(* IEC 61131-3 sources: daoli-st-library/DL_MathData (part 6) *)

(* ---- FC_DL_StringToUdintEx.st ---- *)
(*
    组件名称 : FC_DL_StringToUdintEx
    所属子库 : DL_MathData
    当前版本 : 1.0.0
    兼 容 性 : CODESYS V3.5+ / TwinCAT 3 / 汇川 InoProShop；仅依赖 Standard.library
    溯源声明 : IEC 61131-3 标准语义的道莅防御性实现
              （解析口径复用库内 FC_DL_StringToDint 的四态状态机与判界结构，
                按无符号域重写判界；零外部源码复制，参考实现仅限 MIT/Apache 许可）
    功能描述 : 无符号整数字符串严格解析（UDINT 域，配方号 / 计数器预置 / 批次号）。
              取舍 ①：不委托任何平台串转数值内建——三家平台对非法字符、前导空格、
              符号重复的处理各不相同，有的返回 0、有的抛异常、有的静默截断，且都
              不告诉调用方错在第几位；本件逐字符推进，判断口径完全一致，并给出
              首个非法字符位置。
              取舍 ②：空格一律按非法字符拒绝（与 FC_DL_StringToDint 的「忽略空格
              并提示」口径刻意分叉）——UDINT 域多为机器写入值，隐式吞空格易掩盖
              脏数据，从严拒绝并在 nErrPos 定位。
              取舍 ③：升位到 LINT 累加，每步先判界再落账——UDINT 域中间量在
              429496729 × 10 + 5 处已越界，直接在 UDINT/DINT 里累加必然回绕
              （R241 口径：跨类型降型禁靠隐式回绕兜底）；LINT 域足够宽，判界
              判的是 LINT 与 UDINT 上界的比较，安全。
              取舍 ④：溢出后返回「夹到上界」的值并置 bValid = FALSE——夹域值便于
              现场看出「方向对了但超了」；同时绝不把夹域值当有效值输出。
              取舍 ⑤：负号一律判越域拒绝（含 −0）——UDINT 无负域，负号属语义错误
              而非语法错误，独立占码与非法字符区分。
    本文件内含 : FUNCTION FC_DL_StringToUdintEx（单 POU）
                 同文件 TYPE E_DL_StrToUdintState（归属本函数，全库唯一）
    依 赖    : 无 DL_ 内部依赖；Standard.library: LEN / MID / FIND
    错误码   : 16#0001_03D6 [故障级] 空串或仅符号，nErrPos = 长度 + 1，返回 0，bValid = FALSE
               16#0001_03D7 [故障级] 负值越 UDINT 域（含 −0，从严拒绝），返回 0，bValid = FALSE
               16#0001_03D8 [故障级] 数值溢出，返回夹到上界的值，bValid = FALSE
               16#0001_03D9 [故障级] 非法字符（含 CASE 落 ELSE 的非法状态兜底与扫描失控复用，
                             不新占码位），返回 0，bValid = FALSE
               （R90 反证句：四类故障场景的输出组合互不相同——空串与非法字符返回 0、
                 溢出返回上界夹域值、负值返回 0 但 nErrPos 定位在符号位；返回值加
                 nErrPos 无法唯一还原「空串」与「负值」（同为 0），故两场景各自占码）
    红线自检 : R1 ✓ 零全局变量与外部变量 ｜ R2 ✓ 零物理 IO 地址
              R3 ✓ 纯 IEC 61131-3 ｜ R4 ✓ 空串闸 + 非法字符定位 + 先判界后落账 + WHILE 守卫计数器
              R5 ✓ 全变量中英双语同行注释 ｜ R6 ✓ ENUM + CASE + ELSE 兜底（非法状态复用 03D9）
              R7 N/A 无定时器、无沿检测实例 ｜ R8 ✓ 上下界、长度上限、守卫上限全常量化
    修订历史 :
        2026-11-19  v1.0.0  首版，R40 批次 3 入库
*)

(*-----------------------------------------------------------------------------
 * 枚举: E_DL_StrToUdintState（归属本函数，与其同文件发布，全库唯一）
 * 含义: 逐字符解析的四态推进，成员值写死便于工程持久化
 *----------------------------------------------------------------------------*)
TYPE E_DL_StrToUdintState :
(
    eLeadSpace := 0,    // 起始态：空格按非法字符拒绝，遇其余字符转符号态 ｜ start state, blanks are rejected as illegal, any other character moves to the sign state
    eSign      := 10,   // 符号态：取前导 +/− 号或直接进数字态 ｜ sign state, consumes the leading sign or falls through to the digits
    eDigits    := 20,   // 数字态：逐位累加，遇非数字一律非法 ｜ digits state, accumulates digit by digit, any non-digit is illegal
    eDone      := 30    // 结束态：串尾守卫态，任何字符均非法 ｜ done state, an end-of-string guard, any character here is illegal
);
END_TYPE

FUNCTION FC_DL_StringToUdintEx : UDINT
VAR_INPUT
    sIn             : STRING;           // 待解析文本，最长 255 字符，不允许任何空格 [字符] ｜ input text, up to 255 characters, no blanks allowed [char]
    bAllowSign      : BOOL := FALSE;    // 是否允许前导 +/− 号，UDINT 口径缺省禁止 ｜ whether a leading sign is allowed, the UDINT mode forbids it by default
END_VAR
VAR_OUTPUT
    eErr            : UDINT;           // 错误码，0=正常；16#0001_03XX 故障级 ｜ error id, 0=ok, 16#0001_03XX=fault level
    bError          : BOOL;            // 故障级标志，eErr 落 16#0001_03XX 时为 TRUE ｜ fault flag, TRUE on fault-level eErr
    bValid          : BOOL;            // 返回值是否可用 ｜ result usable flag
    nErrPos         : INT;             // 首个非法字符位置（1 基），0 = 无错 [字符] ｜ position of the first illegal character, 1 based, zero means no error [char]
END_VAR
VAR
    eState          : E_DL_StrToUdintState;  // 解析状态机当前态 ｜ current parse state
    nLen            : INT;             // 文本长度，入口锁存一次，其后全部取自该副本 [字符] ｜ latched text length, every later bound comes from this copy [char]
    nPos            : INT;             // 字符游标（1 基）[字符] ｜ character cursor, 1 based [char]
    nGuard          : DINT;            // WHILE 防死锁守卫计数 [次] ｜ loop guard counter [count]
    nDigitVal       : INT;             // 当前字符的数字值，未命中为 −1 [无量纲] ｜ numeric value of the current character, minus one when not a digit [dimensionless]
    nDigits         : INT;             // 已接受的有效数字位数 [位] ｜ number of accepted digits [digit]
    sChar           : STRING(1);       // 当前字符，由标准 MID 取出 [字符] ｜ current character read with the standard MID [char]
    bNeg            : BOOL;            // 负号标志，由前导符号决定 ｜ negative flag set by the leading sign
    bAbort          : BOOL;            // 中止标志，置位后立即退出扫描 ｜ abort flag, the scan stops as soon as it is set
    bOverflow       : BOOL;            // 溢出标志 ｜ overflow flag
    liAcc           : LINT;            // 升位累加器 [无量纲] ｜ widened accumulator [dimensionless]
    liNext          : LINT;            // 下一拍候选累加值，先判界再落账 [无量纲] ｜ candidate accumulator tested before it is committed [dimensionless]
END_VAR
VAR CONSTANT
    DL_UDINT_MAX_LI    : LINT := 4294967295;     // UDINT 上界的 LINT 判界值 [无量纲] ｜ UDINT upper bound as the LINT test limit [dimensionless]
    DL_LINT_TEN        : LINT := 10;             // 十进制进位基数 [无量纲] ｜ decimal radix [dimensionless]
    DL_STR_MAXLEN      : INT := 255;             // 文本长度上限 [字符] ｜ text length upper bound [char]
    DL_STR_GUARD_MAX   : DINT := 600;            // 守卫上限，须大于 255 + 2 次不推进状态 ｜ guard limit, larger than the length plus two non advancing states
    DL_STR_ONE         : INT := 1;               // 单位哨兵 [无量纲] ｜ unity sentinel [dimensionless]
    DL_STR_DIGITS      : STRING := '0123456789'; // 数字字符表，FIND 命中位置 − 1 即数字值 [字符] ｜ digit table, the FIND position minus one is the value [char]
    DL_ERR_NONE        : UDINT := 16#0000_0000;  // 无故障 ｜ no error
END_VAR

// 段 1｜返回值与错误状态预置 ｜ segment 1, preset the return value and the error state
FC_DL_StringToUdintEx := 0;                   // 故障缺省返回 0 ｜ fault default returns zero
eErr           := DL_ERR_NONE;                // 预置无错误 ｜ preset no error
bError         := FALSE;                      // 预置无故障 ｜ preset no fault
bValid         := FALSE;                      // 预置结果不可用 ｜ preset unusable
nErrPos        := 0;                          // 0 表示无错 ｜ zero means no error
eState         := E_DL_StrToUdintState.eLeadSpace;  // 起始态 ｜ start in the start state
nLen           := LEN(sIn);                   // 长度只锁存一次，禁循环内重复 LEN ｜ latch the length once, never call LEN again in the loop
nPos           := DL_STR_ONE;                 // 游标从 1 开始（MID 为 1 基）｜ the cursor starts at one because MID is one based
nGuard         := 0;                          // 守卫清零 ｜ clear the guard
nDigits        := 0;                          // 有效位数清零 ｜ clear the digit count
nDigitVal      := 0;                          // 数字值清零 ｜ clear the digit value
bNeg           := FALSE;                      // 预置无负号 ｜ preset no negative sign
bAbort         := FALSE;                      // 预置不中止 ｜ preset no abort
bOverflow      := FALSE;                      // 预置无溢出 ｜ preset no overflow
liAcc          := 0;                          // 累加器清零 ｜ clear the accumulator
liNext         := 0;                          // 候选值清零 ｜ clear the candidate
sChar          := '';                         // 字符缓冲清空 ｜ clear the character buffer

// 段 2｜逐字符状态机：四态推进，ELSE 兜底拦非法状态 ｜ segment 2, four state machine with an ELSE backstop
WHILE (nPos <= nLen) AND (NOT bAbort) AND (nGuard <= DL_STR_GUARD_MAX) DO
    sChar := MID(sIn, DL_STR_ONE, nPos);    // 取当前位置的一个字符 ｜ take one character at the current position
    CASE eState OF
        E_DL_StrToUdintState.eLeadSpace :
            // 起始态：空格从严拒绝（取舍 ②），其余字符转符号态 ｜ start state: blanks are strictly rejected, any other character moves to the sign state
            IF sChar = ' ' THEN
                eErr    := 16#0001_03D9;    // 空格按非法字符拒绝（故障级）｜ a blank is rejected as an illegal character
                bError  := TRUE;            // 置故障标志 ｜ raise the fault flag
                nErrPos := nPos;            // 定位到空格位 ｜ point at the blank
                bAbort  := TRUE;            // 中止扫描 ｜ abort the scan
            ELSE
                eState := E_DL_StrToUdintState.eSign;  // 转符号态，本拍不消费字符，下一轮重取同一字符 ｜ move to the sign state without consuming this character
            END_IF

        E_DL_StrToUdintState.eSign :
            IF (sChar = '+') OR (sChar = '-') THEN
                IF NOT bAllowSign THEN
                    eErr   := 16#0001_03D9;     // 不允许符号却出现符号（故障级）｜ a sign appeared although it is forbidden
                    bError := TRUE;             // 置故障标志 ｜ raise the fault flag
                    nErrPos := nPos;            // 定位到符号位 ｜ point at the sign
                    bAbort := TRUE;             // 中止扫描 ｜ abort the scan
                ELSE
                    bNeg   := (sChar = '-');    // 负号判定（取舍 ⑤：负号在出口判越域）｜ detect the minus sign (rejected as out-of-domain at the exit)
                    nPos   := nPos + DL_STR_ONE;   // 消费符号 ｜ consume the sign
                    eState := E_DL_StrToUdintState.eDigits;  // 转数字态 ｜ move to the digit state
                END_IF
            ELSE
                eState := E_DL_StrToUdintState.eDigits;  // 无符号直接进数字态 ｜ no sign, go straight to the digits
            END_IF

        E_DL_StrToUdintState.eDigits :
            // 数字态：数字先判界后落账，非数字一律非法（空格含在内，从严口径）｜ digit state: digits are tested before commit, any non-digit is illegal (blanks included, strict mode)
            nDigitVal := FIND(DL_STR_DIGITS, sChar) - DL_STR_ONE;   // 命中 0~9，未命中 −1 ｜ zero to nine when found, minus one otherwise
            IF nDigitVal < 0 THEN
                eErr    := 16#0001_03D9;            // 非法字符（故障级）｜ illegal character, fault level
                bError  := TRUE;                    // 置故障标志 ｜ raise the fault flag
                nErrPos := nPos;                    // 定位到首个非法字符 ｜ point at the first illegal character
                bAbort  := TRUE;                    // 中止扫描 ｜ abort the scan
            ELSE
                liNext := liAcc * DL_LINT_TEN + INT_TO_LINT(nDigitVal);   // 先算候选值 ｜ compute the candidate first
                IF liNext > DL_UDINT_MAX_LI THEN
                    bOverflow := TRUE;              // 越界即溢出，不落账 ｜ beyond the limit means overflow, not committed
                    nErrPos   := nPos;              // 溢出位也必须定位，否则 nErrPos = 0 会被读成「无错」｜ locate the overflowing digit, zero would read as no error
                    bAbort    := TRUE;              // 中止扫描 ｜ abort the scan
                ELSE
                    liAcc   := liNext;              // 落账 ｜ commit
                    nDigits := nDigits + DL_STR_ONE;   // 有效位加一 ｜ one more digit accepted
                    nPos    := nPos + DL_STR_ONE;   // 前进一格 ｜ advance one position
                END_IF
                IF nPos > nLen THEN
                    eState := E_DL_StrToUdintState.eDone;   // 已到串尾，转结束态守卫 ｜ reached the end, move to the done guard
                END_IF
            END_IF

        E_DL_StrToUdintState.eDone :
            // 结束态：本件从严口径，任何尾随字符（含空格）均非法 ｜ done state: in strict mode any trailing character (blanks included) is illegal
            eErr    := 16#0001_03D9;                // 尾随非法字符（故障级）｜ illegal trailing character, fault level
            bError  := TRUE;                        // 置故障标志 ｜ raise the fault flag
            nErrPos := nPos;                        // 定位 ｜ point at the position
            bAbort  := TRUE;                        // 中止扫描 ｜ abort the scan

    ELSE
        // 非法状态兜底：枚举被外部改写或内存损伤，一律按「输入不可解析」处置（R90：复用非法字符码，不新占码位）
        eState   := E_DL_StrToUdintState.eDone;          // 强制回已知态 ｜ force back to a known state
        eErr     := 16#0001_03D9;                        // 复用非法字符码 ｜ reuse the illegal character code
        bError   := TRUE;                               // 置故障标志 ｜ raise the fault flag
        nErrPos  := nPos;                               // 定位当前位 ｜ point at the current position
        bAbort   := TRUE;                               // 中止扫描 ｜ abort the scan
    END_CASE
    nGuard := nGuard + 1;                              // 守卫递增 ｜ increment the guard
END_WHILE

// 段 3｜守卫复检：理论不可达（长度 ≤ 255，不推进状态最多 2 次）｜ segment 3, guard re-check, unreachable in theory
IF nGuard > DL_STR_GUARD_MAX THEN
    FC_DL_StringToUdintEx := 0;        // 不给可疑结果 ｜ never emit a suspicious result
    eErr   := 16#0001_03D9;            // 扫描失控复用非法字符码（不新占码位）｜ a runaway scan reuses the illegal character code
    bError := TRUE;                    // 置故障标志 ｜ raise the fault flag
    nErrPos := nPos;                   // 定位 ｜ point at the current position
    RETURN;                            // bValid 保持 FALSE ｜ bValid stays FALSE
END_IF

// 段 4｜非法/溢出已中止：直接出口（故障行为已在扫描中定性）｜ segment 4, exit when the scan was aborted
IF bAbort THEN
    IF bOverflow THEN
        FC_DL_StringToUdintEx := 4294967295; // 溢出夹到 UDINT 上界 ｜ overflow saturated to the UDINT upper bound
        eErr := 16#0001_03D8;        // 溢出已夹上界（故障级）｜ overflow saturated, fault level
        bError := TRUE;              // 置故障标志（R45 配对，扫描内溢出只置 bOverflow，出口统一配对）｜ raise the fault flag (R45 pairing)
    ELSE
        FC_DL_StringToUdintEx := 0;  // 语法错误返回 0 ｜ a syntax error returns zero
    END_IF
    RETURN;                          // bValid 保持 FALSE ｜ bValid stays FALSE
END_IF

// 段 5｜空串或仅符号闸 ｜ segment 5, empty string or sign-only gate
IF nDigits = 0 THEN
    FC_DL_StringToUdintEx := 0;         // 无有效数字返回 0 ｜ no digit at all, return zero
    eErr    := 16#0001_03D6;            // 空串或仅符号（故障级）｜ empty or sign only, fault level
    bError  := TRUE;                    // 置故障标志（R45 配对）｜ raise the fault flag (R45 pairing)
    nErrPos := nLen + DL_STR_ONE;       // 指向「串尾后一位」，与库内同族口径一致 ｜ point past the end, consistent with the sibling component
    RETURN;                             // bValid 保持 FALSE ｜ bValid stays FALSE
END_IF

// 段 6｜负值越域闸（取舍 ⑤：负号含 −0 一律从严拒绝）｜ segment 6, negative out-of-domain gate (a minus sign including minus zero is strictly rejected)
IF bNeg THEN
    FC_DL_StringToUdintEx := 0;         // 负值越域返回 0 ｜ out-of-domain negative returns zero
    eErr    := 16#0001_03D7;            // 负值越 UDINT 域（故障级）｜ negative beyond the UDINT domain, fault level
    bError  := TRUE;                    // 置故障标志（R45 配对）｜ raise the fault flag (R45 pairing)
    nErrPos := DL_STR_ONE;              // 定位到符号位（第 1 位）｜ point at the sign position (position one)
    RETURN;                             // bValid 保持 FALSE ｜ bValid stays FALSE
END_IF

// 段 7｜出口装配：累加器域内单点落账 ｜ segment 7, exit assembly: the accumulator is in-domain, commit once
FC_DL_StringToUdintEx := LINT_TO_UDINT(liAcc); // 判界已保证 liAcc ≤ UDINT 上界，降型安全 ｜ the domain test guarantees the accumulator is within the UDINT bound, the down-conversion is safe
bValid := TRUE;                      // 结果可用 ｜ the result is usable
END_FUNCTION

(* ---- FC_DL_SwapBytes32.st ---- *)
(*==============================================================================
 * 组件名称 (Component)  : FC_DL_SwapBytes32
 * 所属子库 (Sublibrary) : DL_MathData
 * 当前版本 (Version)    : 1.0.0
 * 兼容性   (Platform)   : CODESYS 3.5 / TwinCAT 3 / 汇川 InoProShop / Machine Expert
 *                         仅依赖 Standard.library 的 SHL / SHR / AND / OR，零厂商方言
 * 功能描述 (Function)   : 32 位量四排布（ABCD / DCBA / BADC / CDAB）归一化转换。
 *                         调用方声明通信侧原始拼接值实际所属的排布，
 *                         函数统一输出 ABCD（大端大字）归一化值。
 *                         语义锁定为单向归一化，不做双向目标排布选择；
 *                         需要反向时以对称排布重新声明即可（四排布两两互逆）。
 *                         用于 Modbus 多寄存器浮点/长整型量"读回 1e38 天文数字"的定位与校正。
 * 开源溯源 (Origin)     : 原创实现。四种排布命名与业界别名（字交换 / 寄存器内字节互换 /
 *                         全反序）参照 modbus.org 公开协议说明与多家转换器技术资料的
 *                         事实约定；本文件为独立重构，未复制任何源码。
 * 本文件内含       : TYPE  E_DL_ByteOrder（配套枚举，归属 DL_MathData）
 *                    FC    FC_DL_SwapBytes32
 * 依赖     (Depends)    : 无 DL_ 内部依赖；Standard.library: SHL / SHR
 * 红线自检 (Redline)    : R1 ✓ 禁用全局存储与物理寻址 ｜ R2 ✓ 无地址直写
 *                         R3 ✓ 移位掩码提取 + 显式类型转换，无切片/指针/字节方言
 *                         R4 N/A（无除法/数组/循环/浮点）｜ R5 ✓ 全变量中英双语同行注释
 *                         R6 ✓ 四排布 CASE 分派 + ELSE 兜底 ｜ R7 N/A（无定时器/边沿实例）
 *                         R8 ✓ 移位量与掩码全常量化
 *
 * 【实现选择 / Implementation choice（边界 B6）】
 *   四条转换路径全部用"移位提取 + 显式 BYTE 转换 + 移位重装"实现，
 *   不调用 16 位互换构件，保证本文件自洽、可单独编译与单独单测。
 *
 * 【浮点使用口径 / Float usage（边界 B7）】
 *   本函数只输出归一化 DWORD，不做 DWORD 到 REAL 的二进制重解释。
 *   浮点拼接规则各平台存在差异，由调用方按其平台口径完成，避免在本层引入行为分支。
 *
 * 【验收向量 / Acceptance vectors（边界 B5，已复算）】
 *   以 16#12345678 为基准：ABCD → 16#12345678；DCBA → 16#78563412；
 *   BADC → 16#34127856；CDAB → 16#56781234。
 *
 * 修订历史 (Revision)   :
 *   2026-11-14  v1.0.0  首版入库（Phase 1 第二轮 · Level 0 批次 C）
 *============================================================================*)

(*-----------------------------------------------------------------------------
 * 枚举: E_DL_ByteOrder（归属 DL_MathData，与 FC_DL_SwapBytes32 同文件）
 * 含义: 通信侧 32 位量的字节排布。A 为最高字节（位 31..24），D 为最低字节。
 *----------------------------------------------------------------------------*)
TYPE E_DL_ByteOrder :
(
    eAbcd := 0,    // ABCD：大端大字（Modicon 事实标准），原始值无需转换 / Big-endian big-word, pass-through
    eDcba := 1,    // DCBA：四字节全反序，常见于小端 CPU 直出的协议栈 / Full byte reverse
    eBadc := 2,    // BADC：两个寄存器内部各自字节互换 / Byte swap within each register
    eCdab := 3     // CDAB：高低字交换（寄存器字序反），常见于电能表 / Word swap
);
END_TYPE

FUNCTION FC_DL_SwapBytes32 : DWORD
VAR_INPUT
    uRaw      : DWORD;                        // 通信侧原始 32 位拼接值 / Raw 32-bit value assembled from comms
    eRawOrder : E_DL_ByteOrder := eAbcd;      // 声明原始值所属排布 / Declared byte order of raw value
END_VAR
VAR_OUTPUT
    bValid    : BOOL;                         // 排布枚举合法标志 / Order enum valid flag
    uErrorId  : UDINT;                        // 故障码，0 = 无故障 / Error code, 0 = no error
END_VAR
VAR
    uA : BYTE;   // 字节 A（uRaw 位 31..24） / Byte A, bits 31..24
    uB : BYTE;   // 字节 B（uRaw 位 23..16） / Byte B, bits 23..16
    uC : BYTE;   // 字节 C（uRaw 位 15..8）  / Byte C, bits 15..8
    uD : BYTE;   // 字节 D（uRaw 位 7..0）   / Byte D, bits 7..0
END_VAR
VAR CONSTANT
    DL_SWAP_SHIFT8  : UDINT := 8;               // 字节移位量 [bit] / Byte shift width [bit]
    DL_SWAP_SHIFT16 : UDINT := 16;              // 字移位量 [bit] / Word shift width [bit]
    DL_SWAP_SHIFT24 : UDINT := 24;              // 最高字节移位量 [bit] / Top byte shift width [bit]
    DL_MASK_BYTE    : DWORD := 16#0000_00FF;    // 单字节掩码 / Single-byte mask
END_VAR

(*------------------------------------------------------------------------------
 * 段 1｜安全预置（边界 B1 / P-01）：先返回原值，任何异常路径都不会返回 0
 *      Safe preset: return the raw value first, no exceptional path returns zero
 *      0 对浮点量是合法灾难值，原值直通是最安全的确定值
 *      Zero is a legal but catastrophic float value, pass-through is the safest result
 *-----------------------------------------------------------------------------*)
FC_DL_SwapBytes32 := uRaw;
bValid   := TRUE;
uErrorId := 16#0000_0000;

(*------------------------------------------------------------------------------
 * 段 2｜字节提取（边界 B2）：仅移位 + 掩码 + 显式 BYTE 转换，禁止切片与指针
 *      Byte extraction: shift + mask + explicit BYTE conversion only
 *-----------------------------------------------------------------------------*)
uA := DWORD_TO_BYTE(SHR(uRaw, DL_SWAP_SHIFT24) AND DL_MASK_BYTE);
uB := DWORD_TO_BYTE(SHR(uRaw, DL_SWAP_SHIFT16) AND DL_MASK_BYTE);
uC := DWORD_TO_BYTE(SHR(uRaw, DL_SWAP_SHIFT8)  AND DL_MASK_BYTE);
uD := DWORD_TO_BYTE(uRaw AND DL_MASK_BYTE);

(*------------------------------------------------------------------------------
 * 段 3｜四排布分派（边界 B3/B4）：CASE 分派禁止 IF 链，ELSE 兜底拒收非法枚举
 *      Four-order dispatch: CASE only, ELSE intercepts an out-of-domain enum
 *-----------------------------------------------------------------------------*)
CASE eRawOrder OF

    eAbcd:
        (* 大端大字已是归一化目标，原值直通 *)
        (* Big-endian big-word is already the normalised target, pass through *)
        FC_DL_SwapBytes32 := uRaw;

    eDcba:
        (* 全反序：D C B A *)
        (* Full byte reverse: D C B A *)
        FC_DL_SwapBytes32 := (SHL(BYTE_TO_DWORD(uD), DL_SWAP_SHIFT24)
                          OR  SHL(BYTE_TO_DWORD(uC), DL_SWAP_SHIFT16)
                          OR  SHL(BYTE_TO_DWORD(uB), DL_SWAP_SHIFT8)
                          OR  BYTE_TO_DWORD(uA));

    eBadc:
        (* 寄存器内字节互换：B A D C *)
        (* Byte swap within each register: B A D C *)
        FC_DL_SwapBytes32 := (SHL(BYTE_TO_DWORD(uB), DL_SWAP_SHIFT24)
                          OR  SHL(BYTE_TO_DWORD(uA), DL_SWAP_SHIFT16)
                          OR  SHL(BYTE_TO_DWORD(uD), DL_SWAP_SHIFT8)
                          OR  BYTE_TO_DWORD(uC));

    eCdab:
        (* 高低字交换：C D A B *)
        (* Word swap: C D A B *)
        FC_DL_SwapBytes32 := (SHL(BYTE_TO_DWORD(uC), DL_SWAP_SHIFT24)
                          OR  SHL(BYTE_TO_DWORD(uD), DL_SWAP_SHIFT16)
                          OR  SHL(BYTE_TO_DWORD(uA), DL_SWAP_SHIFT8)
                          OR  BYTE_TO_DWORD(uB));

    ELSE
        (* 非法枚举拦截：枚举被强制写入定义域外的值时返回原值并报错 *)
        (* Illegal enum interception: keep the raw value and raise the error *)
        FC_DL_SwapBytes32 := uRaw;
        bValid            := FALSE;
        uErrorId          := 16#0001_000E;

END_CASE;
END_FUNCTION

(* ---- FC_DL_TableIndexBinarySearch.st ---- *)
(*==============================================================================
 * 组件名称 (Component)  : FC_DL_TableIndexBinarySearch
 * 所属子库 (Sublibrary) : DL_MathData
 * 当前版本 (Version)    : 1.0.0
 * 兼容性   (Platform)   : CODESYS 3.5+ / TwinCAT 3 / 汇川 InoProShop / 施耐德 Machine Expert
 *                         仅依赖 IEC 61131-3 标准数学（ABS / MIN / MAX），零厂商私有库
 * 功能描述 (Function)   : **升序**节点表二分查找定位（O(log n)），返回区间左端下标与段内比例。
 *                         迭代式二分：维护 [iLo, iHi] 使 afX[iLo] <= fXin <= afX[iHi]，
 *                         每次收缩一半，直到 iHi - iLo = 1，此时 iSeg = iLo。
 *                         32 点表最多 5 次迭代（2^5 = 32），循环上界显式封顶 8 次，
 *                         结构上不可能死循环（R6 周期安全：纯函数虽无跨周期状态，
 *                         仍对不可终止循环做硬保护）。
 *                         用途：大表（温压补偿、阀门口径选型）的高频查表，替代线性扫描。
 * 接口     (Interface)  : 输入 afX 升序节点表 [任意工程量]、iCount 有效点数 [个]（2..32）、
 *                         fXin 查询点 [同 afX 单位]；
 *                         输出 iSeg 区间左端下标 [1..iCount-1]、fRatio 段内比例 [0..1]、
 *                         bExact 是否恰命中节点、bClamped 越界钳位回执、
 *                         eErrCode（E_DL_TblBsearchErr）；
 *                         返回值 = bValid 定位可信标志（TRUE = iSeg/fRatio 可信）。
 * 边界     (Boundary)   : ① 属主边界：只做定位，不做取值；表必须升序（降序表用
 *                         FC_DL_TableLookupDescending）。
 *                         ② 点数域闸 2..32；越域 → 故障级 eBadCount。
 *                         ③ 非有限双判：查询点 + 全部表元素逐项枚举（漏判单个元素会使比较静默失效）。
 *                         ④ 升序性校验：二分不校验全序，但会校验命中区间的两个端点是否满足
 *                         afX[iSeg] <= afX[iSeg+1]，违反即判 eTableNotAsc（防止强序假设）。
 *                         ⑤ 段宽近似零 → fRatio 置 0 并置信息级 eDegenerateSeg（除零防护）。
 *                         ⑥ 迭代次数硬上界 DL_TBC_ITER_MAX = 8，超出即判 eSearchOverflow
 *                         （理论上不可达，作为不可终止循环的兜底闸）。
 *                         ⑦ 零全局耦合（无 GVL / VAR_EXTERNAL / 物理地址）。
 * 分工声明 (Scope)      : 与 `FC_DL_TableLookupDescending` 分工：降序 / 线性归那件、
 *                         升序 / 二分归本件；与 `FC_DL_InterpSegmentWeight` 分工：
 *                         权重归那件、本件只给下标与比例。
 * 来源标签 (Source Tag) : 原创实现（无外部代码引入）
 * 码表     (Codes)      : 本件不占用全局数字码位；出口为 BOOL + INT + LREAL + 2×BOOL +
 *                         本文件内定义 enum E_DL_TblBsearchErr（全库唯一）。
 * 红线自检 (Redline)    : R1 ✓ 零 GVL/VAR_EXTERNAL ｜ R2 ✓ 零 %I/%Q/%M ｜ R3 ✓ 纯 IEC 61131-3
 *                         R4 ✓ 点数域闸 + 全表非有限双判 + 段宽判零 + 迭代次数硬上界 ｜ R5 ✓ 声明逐行同行双语注释
 *                         R6 N/A（纯函数无状态机；循环不可终止风险由迭代上限拦截） ｜ R7 N/A（无实例调用）
 * 修订历史 (Revision)   : 2026-11-23  v1.0.0  R77 首版（批次 B3 · 序号 5）
 * 验收向量 (Acceptance) : ① afX=[0,10,20,30], iCount=4, fXin=15 → iSeg=2,
 *                         fRatio=(15-10)/(20-10)=0.5, bExact=FALSE, bClamped=FALSE, eOk；
 *                         ② afX 同上, fXin=20 → iSeg=2（恰命中右端）, bExact=TRUE；
 *                         ③ afX 同上, fXin=-5 → iSeg=1, fRatio=0.0, bClamped=TRUE, eOk；
 *                         ④ afX 同上, fXin=100 → iSeg=3, fRatio=1.0, bClamped=TRUE, eOk；
 *                         ⑤ iCount=40 → 返回 FALSE, iSeg=0, eBadCount。
 *==============================================================================*)

(*-----------------------------------------------------------------------------
 * 枚举: E_DL_TblBsearchErr（升序表二分查找错误码，归属 DL_MathData，与本件同文件，全库唯一属主）
 *----------------------------------------------------------------------------*)
TYPE E_DL_TblBsearchErr :
(
    eOk              := 0,   // 信息级：定位完成 / Info: located
    eDegenerateSeg   := 1,   // 信息级：段宽近似零，比例置 0 / Info: degenerate segment, ratio zeroed
    eBadCount        := 2,   // 故障级：点数越域 / Fault: point count out of domain
    eNonFinite       := 3,   // 故障级：查询点或表元素非有限 / Fault: query or table entry non-finite
    eTableNotAsc     := 4,   // 故障级：表不满足升序约定 / Fault: table violates ascending contract
    eSearchOverflow  := 5    // 故障级：迭代超上限（不可达兜底） / Fault: iteration overflow, unreachable guard
);
END_TYPE

FUNCTION FC_DL_TableIndexBinarySearch : BOOL
VAR_INPUT
    afX    : ARRAY[1..32] OF LREAL;  // 升序节点表 [任意工程量] / Ascending node table
    iCount : INT;                    // 有效点数（2..32） [个] / Valid point count, 2..32
    fXin   : LREAL;                  // 查询点 [同 afX 单位] / Query value
END_VAR
VAR_OUTPUT
    iSeg     : INT;    // 区间左端下标（1..iCount-1） [-] / Segment left index
    fRatio   : LREAL;  // 段内比例（0 = 左端，1 = 右端） [-] / In-segment ratio
    bExact   : BOOL;   // 是否恰命中节点 [-] / Whether a node was hit exactly
    bClamped : BOOL;   // 越界钳位回执 [-] / Out-of-range clamp receipt
    eErrCode : E_DL_TblBsearchErr; // 错误码出口 [-] / Error code outlet
END_VAR
VAR
    _i       : INT;    // 表元素遍历下标 [-] / Table traversal index
    _iLo     : INT;    // 二分下界 [-] / Binary search low bound
    _iHi     : INT;    // 二分上界 [-] / Binary search high bound
    _iMid    : INT;    // 二分中点 [-] / Binary search midpoint
    _iIter   : INT;    // 迭代计数 [-] / Iteration counter
    _bNonFin : BOOL;   // 非有限标志 [-] / Non-finite flag
    _fDen    : LREAL;  // 段宽（分母） [-] / Segment width denominator
    _fRatio  : LREAL;  // 未钳位比例 [-] / Raw ratio
END_VAR
VAR CONSTANT
    DL_TBC_CNT_MIN  : INT := 2;        // 点数下限 [个] / Count lower bound
    DL_TBC_CNT_MAX  : INT := 32;       // 点数上限（数组容量） [个] / Count upper bound
    DL_TBC_ITER_MAX : INT := 8;        // 迭代次数硬上界（2^8 > 32） [次] / Hard iteration bound
    DL_TBC_TINY     : LREAL := 1.0E-9; // 段宽与命中近似零阈值 [-] / Degenerate and exact threshold
    DL_TBC_ZERO     : LREAL := 0.0;    // 零与比例下限 [-] / Zero and ratio lower bound
    DL_TBC_ONE      : LREAL := 1.0;    // 比例上限 [-] / Ratio upper bound
    DL_TBC_HALF     : INT := 2;        // 二分除数（整数除） [-] / Binary divisor, integer division
END_VAR

(* —— 段 0：出口预置安全值 —— *)
FC_DL_TableIndexBinarySearch := FALSE;             // 返回值预置无效 / Return preset invalid
iSeg     := 0;                                     // 下标哨兵 / Index sentinel
fRatio   := DL_TBC_ZERO;                           // 比例哨兵 / Ratio sentinel
bExact   := FALSE;                                 // 恰命中标志预置否 / Exact flag preset false
bClamped := FALSE;                                 // 钳位回执预置否 / Clamp receipt preset false
eErrCode := E_DL_TblBsearchErr.eBadCount;          // 预置最严码 / Preset strictest code

(* —— 段 1：点数域闸 —— *)
IF (iCount < DL_TBC_CNT_MIN) OR (iCount > DL_TBC_CNT_MAX) THEN
    RETURN;
END_IF

(* —— 段 2：非有限域闸（查询点 + 全部表元素逐项枚举） —— *)
_bNonFin := (fXin <> fXin) OR ((fXin - fXin) <> DL_TBC_ZERO);
_i := 1;
WHILE _i <= iCount DO
    IF (afX[_i] <> afX[_i]) OR ((afX[_i] - afX[_i]) <> DL_TBC_ZERO) THEN
        _bNonFin := TRUE;
    END_IF
    _i := _i + 1;
END_WHILE
IF _bNonFin THEN
    eErrCode := E_DL_TblBsearchErr.eNonFinite;
    RETURN;
END_IF

(* —— 段 3：上下越界早退（钳到端段，避免二分越出下标域） —— *)
IF fXin <= afX[1] THEN
    iSeg     := 1;
    fRatio   := DL_TBC_ZERO;
    bClamped := TRUE;
    bExact   := (ABS(afX[1] - fXin) < DL_TBC_TINY);   // 恰落在首节点 / Exactly on first node
    eErrCode := E_DL_TblBsearchErr.eOk;
    FC_DL_TableIndexBinarySearch := TRUE;
    RETURN;
END_IF
IF fXin >= afX[iCount] THEN
    iSeg     := iCount - 1;
    fRatio   := DL_TBC_ONE;
    bClamped := TRUE;
    bExact   := (ABS(afX[iCount] - fXin) < DL_TBC_TINY);   // 恰落在末节点 / Exactly on last node
    eErrCode := E_DL_TblBsearchErr.eOk;
    FC_DL_TableIndexBinarySearch := TRUE;
    RETURN;
END_IF

(* —— 段 4：迭代式二分收缩（迭代次数硬上界，不可终止即兜底判错） —— *)
_iLo   := 1;
_iHi   := iCount;
_iIter := 0;
WHILE ((_iHi - _iLo) > 1) AND (_iIter < DL_TBC_ITER_MAX) DO
    _iMid := (_iLo + _iHi) / DL_TBC_HALF;          // 整数除取中点 / Integer midpoint
    IF fXin >= afX[_iMid] THEN
        _iLo := _iMid;                             // 抬下界 / Raise low bound
    ELSE
        _iHi := _iMid;                             // 压下界 / Lower high bound
    END_IF
    _iIter := _iIter + 1;
END_WHILE

IF (_iHi - _iLo) > 1 THEN
    eErrCode := E_DL_TblBsearchErr.eSearchOverflow; // 迭代未收敛：兜底判错 / Not converged: guard fault
    RETURN;
END_IF

(* —— 段 5：区间端点升序校验（防止强序假设静默失效） —— *)
IF afX[_iLo + 1] < afX[_iLo] THEN
    eErrCode := E_DL_TblBsearchErr.eTableNotAsc;   // 表不满足升序 / Table violates ascending contract
    RETURN;
END_IF

(* —— 段 6：段内比例计算（段宽判零） —— *)
_fDen := afX[_iLo + 1] - afX[_iLo];                // 升序段宽恒 >= 0 / Ascending segment width
IF ABS(_fDen) < DL_TBC_TINY THEN
    fRatio   := DL_TBC_ZERO;                       // 退化段：比例置 0 / Degenerate: ratio zero
    eErrCode := E_DL_TblBsearchErr.eDegenerateSeg; // 信息级码 / Info code
ELSE
    _fRatio  := (fXin - afX[_iLo]) / _fDen;        // 标准比例式 / Standard ratio
    fRatio   := MIN(MAX(_fRatio, DL_TBC_ZERO), DL_TBC_ONE);   // 显式约束 0..1 / Constrain 0..1
    eErrCode := E_DL_TblBsearchErr.eOk;            // 信息级成功 / Info success
END_IF
iSeg := _iLo;                                      // 导出下标 / Export index

(* —— 段 7：恰命中判定（两端节点任一在容差内） —— *)
bExact := (ABS(afX[_iLo] - fXin) < DL_TBC_TINY) OR (ABS(afX[_iLo + 1] - fXin) < DL_TBC_TINY);

(* —— 段 8：下标复检（必须落在 1..iCount-1） —— *)
IF (iSeg < 1) OR (iSeg > (iCount - 1)) THEN
    iSeg     := 0;
    fRatio   := DL_TBC_ZERO;
    bExact   := FALSE;
    eErrCode := E_DL_TblBsearchErr.eTableNotAsc;
    RETURN;
END_IF

FC_DL_TableIndexBinarySearch := TRUE;              // 定位有效 / Lookup valid

END_FUNCTION

(* ---- FC_DL_TableLookupDescending.st ---- *)
(*==============================================================================
 * 组件名称 (Component)  : FC_DL_TableLookupDescending
 * 所属子库 (Sublibrary) : DL_MathData
 * 当前版本 (Version)    : 1.0.0
 * 兼容性   (Platform)   : CODESYS 3.5+ / TwinCAT 3 / 汇川 InoProShop / 施耐德 Machine Expert
 *                         仅依赖 IEC 61131-3 标准数学（ABS / MIN / MAX），零厂商私有库
 * 功能描述 (Function)   : **降序**节点表区间定位（返回区间下标 + 段内比例）。
 *                         适用场景：工艺曲线以「高压→低压」「高温→低温」顺序录入的表格
 *                         （与升序表件互为镜像，避免调用方每次传入前自行反转数组）。
 *                         定位规则：找到 i 使 afX[i] >= fXin >= afX[i+1]，返回
 *                         iSeg = i（区间左端下标）与 fRatio = (afX[i]-fXin)/(afX[i]-afX[i+1])
 *                         （0 = 落在左端节点，1 = 落在右端节点）。
 *                         越界处理：fXin 高于首节点 → iSeg=1、fRatio=0 并置 bClamped；
 *                         fXin 低于末节点 → iSeg=iCount-1、fRatio=1 并置 bClamped
 *                         （钳位语义：不外推，结果恒落在表端点上）。
 * 接口     (Interface)  : 输入 afX 降序节点表 [任意工程量]、iCount 有效点数 [个]（2..32）、
 *                         fXin 查询点 [同 afX 单位]；
 *                         输出 iSeg 区间左端下标 [1..iCount-1]、fRatio 段内比例 [0..1]、
 *                         bClamped 越界钳位回执、eErrCode（E_DL_TblDescErr）；
 *                         返回值 = bValid 定位可信标志（TRUE = iSeg/fRatio 可信）。
 * 边界     (Boundary)   : ① 属主边界：只做定位，不做插值取值（取值归插值族），不修改表。
 *                         ② 点数域闸 2..32；越域 → 故障级 eBadCount。
 *                         ③ 非有限双判：fXin 与**全部参与判据的表元素**（1..iCount）逐个判，
 *                         任一非有限 → 故障级 eNonFinite（漏判单个元素会使距离/比较静默失效）。
 *                         ④ 降序性校验：定位循环未命中即判 eTableNotDesc（表录入违反降序约定），
 *                         不做「假设有序继续算」的静默容错。
 *                         ⑤ 段宽近似零（|afX[i]-afX[i+1]| < 1E-9）→ fRatio 置 0 并置信息级
 *                         eDegenerateSeg（退化段，避免除零；重复节点属录入缺陷需上游修）。
 *                         ⑥ 零全局耦合（无 GVL / VAR_EXTERNAL / 物理地址）。
 * 分工声明 (Scope)      : 与 `FC_DL_TableIndexBinarySearch`（升序 / O(log n)）互为镜像，
 *                         本件为降序线性扫描；与 `FC_DL_InterpSegmentWeight` 分工：
 *                         权重归那件，本件只给下标与比例。
 * 来源标签 (Source Tag) : 原创实现（无外部代码引入）
 * 码表     (Codes)      : 本件不占用全局数字码位；出口为 BOOL + INT + 2×LREAL + BOOL +
 *                         本文件内定义 enum E_DL_TblDescErr（全库唯一）。
 * 红线自检 (Redline)    : R1 ✓ 零 GVL/VAR_EXTERNAL ｜ R2 ✓ 零 %I/%Q/%M ｜ R3 ✓ 纯 IEC 61131-3
 *                         R4 ✓ 点数域闸 + 全表元素非有限双判 + 段宽判零 + 越界钳位 ｜ R5 ✓ 声明逐行同行双语注释
 *                         R6 N/A（纯函数无状态机） ｜ R7 N/A（无实例调用）
 * 修订历史 (Revision)   : 2026-11-23  v1.0.0  R77 首版（批次 B3 · 序号 1）
 * 验收向量 (Acceptance) : ① afX=[100,80,60,40], iCount=4, fXin=90 → 区间 1，
 *                         fRatio=(100-90)/(100-80)=0.5, bClamped=FALSE, eOk；
 *                         ② afX 同上, fXin=110 → iSeg=1, fRatio=0.0, bClamped=TRUE, eOk；
 *                         ③ afX 同上, fXin=10 → iSeg=3, fRatio=1.0, bClamped=TRUE, eOk；
 *                         ④ iCount=1 → 返回 FALSE, iSeg=0, eBadCount；
 *                         ⑤ afX=[100,80,90,40]（非降序）, fXin=85 → 返回 FALSE, eTableNotDesc。
 *==============================================================================*)

(*-----------------------------------------------------------------------------
 * 枚举: E_DL_TblDescErr（降序表定位错误码，归属 DL_MathData，与本件同文件，全库唯一属主）
 *----------------------------------------------------------------------------*)
TYPE E_DL_TblDescErr :
(
    eOk             := 0,   // 信息级：定位完成 / Info: located
    eDegenerateSeg  := 1,   // 信息级：段宽近似零，比例已置 0 / Info: degenerate segment, ratio forced to zero
    eBadCount       := 2,   // 故障级：点数越域 / Fault: point count out of domain
    eNonFinite      := 3,   // 故障级：查询点或表元素非有限 / Fault: query or table entry non-finite
    eTableNotDesc   := 4    // 故障级：表不满足降序约定 / Fault: table violates descending contract
);
END_TYPE

FUNCTION FC_DL_TableLookupDescending : BOOL
VAR_INPUT
    afX    : ARRAY[1..32] OF LREAL;  // 降序节点表 [任意工程量] / Descending node table, any engineering unit
    iCount : INT;                    // 有效点数（2..32） [个] / Valid point count, 2..32
    fXin   : LREAL;                  // 查询点 [同 afX 单位] / Query value, same unit as afX
END_VAR
VAR_OUTPUT
    iSeg     : INT;    // 区间左端下标（1..iCount-1） [-] / Segment left index
    fRatio   : LREAL;  // 段内比例（0 = 左端节点，1 = 右端节点） [-] / In-segment ratio
    bClamped : BOOL;   // 越界钳位回执 [-] / Out-of-range clamp receipt
    eErrCode : E_DL_TblDescErr; // 错误码出口 [-] / Error code outlet
END_VAR
VAR
    _i        : INT;    // 循环下标 [-] / Loop index
    _bFound   : BOOL;   // 区间命中标志 [-] / Segment found flag
    _bNonFin  : BOOL;   // 非有限标志 [-] / Non-finite flag
    _fDen     : LREAL;  // 段宽（分母） [-] / Segment width denominator
    _fRatioIn : LREAL;  // 未钳位比例 [-] / Raw ratio before clamping
END_VAR
VAR CONSTANT
    DL_TDC_CNT_MIN : INT := 2;        // 点数下限 [个] / Count lower bound
    DL_TDC_CNT_MAX : INT := 32;       // 点数上限（数组容量） [个] / Count upper bound, array capacity
    DL_TDC_TINY    : LREAL := 1.0E-9; // 段宽近似零阈值 [-] / Degenerate segment threshold
    DL_TDC_ZERO    : LREAL := 0.0;    // 零与比例下限 [-] / Zero and ratio lower bound
    DL_TDC_ONE     : LREAL := 1.0;    // 比例上限 [-] / Ratio upper bound
END_VAR

(* —— 段 0：出口预置安全值 —— *)
FC_DL_TableLookupDescending := FALSE;              // 返回值预置无效 / Return preset invalid
iSeg     := 0;                                     // 下标哨兵 0（非法下标） / Index sentinel zero
fRatio   := DL_TDC_ZERO;                           // 比例哨兵 0 / Ratio sentinel
bClamped := FALSE;                                 // 钳位回执预置否 / Clamp receipt preset false
eErrCode := E_DL_TblDescErr.eBadCount;             // 预置最严码 / Preset strictest code

(* —— 段 1：点数域闸（数组容量可表性反算） —— *)
IF (iCount < DL_TDC_CNT_MIN) OR (iCount > DL_TDC_CNT_MAX) THEN
    RETURN;                                        // 点数越域：保持故障码与哨兵 / Count out of domain
END_IF

(* —— 段 2：非有限域闸（查询点 + 全部参与判据的表元素逐项枚举） —— *)
_bNonFin := (fXin <> fXin) OR ((fXin - fXin) <> DL_TDC_ZERO);   // 查询点非有限 / Query non-finite
_i := 1;
WHILE _i <= iCount DO
    IF (afX[_i] <> afX[_i]) OR ((afX[_i] - afX[_i]) <> DL_TDC_ZERO) THEN
        _bNonFin := TRUE;                          // 表元素非有限 / Table entry non-finite
    END_IF
    _i := _i + 1;
END_WHILE
IF _bNonFin THEN
    eErrCode := E_DL_TblDescErr.eNonFinite;        // 故障级码 / Fault-level code
    RETURN;
END_IF

(* —— 段 3：上越界钳位（高于首节点：落于首段左端） —— *)
IF fXin >= afX[1] THEN
    iSeg     := 1;
    fRatio   := DL_TDC_ZERO;
    bClamped := TRUE;                              // 钳位回执 / Clamp receipt
    eErrCode := E_DL_TblDescErr.eOk;
    FC_DL_TableLookupDescending := TRUE;
    RETURN;
END_IF

(* —— 段 4：下越界钳位（低于末节点：落于末段右端） —— *)
IF fXin <= afX[iCount] THEN
    iSeg     := iCount - 1;
    fRatio   := DL_TDC_ONE;
    bClamped := TRUE;                              // 钳位回执 / Clamp receipt
    eErrCode := E_DL_TblDescErr.eOk;
    FC_DL_TableLookupDescending := TRUE;
    RETURN;
END_IF

(* —— 段 5：线性扫描定位区间（降序：afX[i] >= fXin >= afX[i+1]） —— *)
_i      := 1;
_bFound := FALSE;
WHILE (_i < iCount) AND (NOT _bFound) DO
    IF (fXin <= afX[_i]) AND (fXin >= afX[_i + 1]) THEN
        _bFound := TRUE;                           // 命中区间 / Segment hit
    ELSE
        _i := _i + 1;                              // 继续右移 / Advance
    END_IF
END_WHILE

IF NOT _bFound THEN
    eErrCode := E_DL_TblDescErr.eTableNotDesc;     // 表不满足降序约定 / Table violates descending contract
    RETURN;                                        // 保持哨兵输出 / Keep sentinel outputs
END_IF

(* —— 段 6：段内比例计算（段宽判零，退化段置 0） —— *)
_fDen := afX[_i] - afX[_i + 1];                    // 降序段宽恒 >= 0 / Descending segment width
IF ABS(_fDen) < DL_TDC_TINY THEN
    fRatio   := DL_TDC_ZERO;                       // 退化段：比例置 0，杜绝除零 / Degenerate: ratio zero, no division
    eErrCode := E_DL_TblDescErr.eDegenerateSeg;    // 信息级码 / Info code
ELSE
    _fRatioIn := (afX[_i] - fXin) / _fDen;         // (左端值 - 查询值) / 段宽 / Ratio formula
    fRatio    := MIN(MAX(_fRatioIn, DL_TDC_ZERO), DL_TDC_ONE);   // 显式约束 0..1 / Constrain into 0..1
    eErrCode  := E_DL_TblDescErr.eOk;              // 信息级成功 / Info success
END_IF
iSeg := _i;                                        // 导出区间左端下标 / Export left index

(* —— 段 7：结果复检（下标必须在 1..iCount-1，比例必须落在 0..1） —— *)
IF (iSeg < 1) OR (iSeg > (iCount - 1)) THEN
    iSeg     := 0;                                 // 下标复检失败回哨兵 / Index recheck failed
    fRatio   := DL_TDC_ZERO;
    eErrCode := E_DL_TblDescErr.eTableNotDesc;     // 保持故障级 / Keep fault-level
    RETURN;
END_IF

FC_DL_TableLookupDescending := TRUE;               // 定位有效 / Lookup valid

END_FUNCTION

(* ---- FC_DL_TableLookupNearestIndex.st ---- *)
(*==============================================================================
 * 组件名称 (Component)  : FC_DL_TableLookupNearestIndex
 * 所属子库 (Sublibrary) : DL_MathData
 * 当前版本 (Version)    : 1.0.0
 * 兼容性   (Platform)   : CODESYS 3.5+ / TwinCAT 3 / 汇川 InoProShop / 施耐德 Machine Expert
 *                         仅依赖 IEC 61131-3 标准数学（ABS），零厂商私有库
 * 功能描述 (Function)   : 最近节点索引查找（等距 / 非等距通用）。遍历 1..iCount 取
 *                         |afX[i] - fXin| 最小者，返回下标与最小距离。
 *                         用途：多档位选型（挡位表 → 最近挡）、配方就近匹配、故障码归类。
 *                         距离采用绝对差（非平方差），仅用于比较与展示，精度足够且无溢出风险。
 *                         并列最小（两节点等距）时保留**较小下标**（首个命中），
 *                         行为确定、可复现，便于验收与回归。
 * 接口     (Interface)  : 输入 afX 节点表（任意升/降序，无需有序） [任意工程量]、
 *                         iCount 有效点数 [个]（1..32）、fXin 查询点 [同 afX 单位]；
 *                         输出 iIndex 最近节点下标 [1..iCount]、fDist 最小绝对距离 [同 afX 单位]、
 *                         eErrCode（E_DL_TblNearErr）；
 *                         返回值 = bValid 查找可信标志（TRUE = iIndex/fDist 可信）。
 * 边界     (Boundary)   : ① 属主边界：只找最近节点，不做插值（插值归插值族）、不要求有序。
 *                         ② 点数域闸 1..32（1 点合法：恒返回该唯一点，距离为其绝对差）。
 *                         ③ 非有限双判：查询点与全部表元素逐个判，任一非有限 → 故障级 eNonFinite。
 *                         ④ 并列最小取较小下标（首个命中即锁定，后续用严格 < 比较），
 *                         保证同输入同输出（无浮点抖动导致的随机化）。
 *                         ⑤ 距离为绝对值，恒非负；复检 distance >= 0 且 < 非有限。
 *                         ⑥ 零全局耦合（无 GVL / VAR_EXTERNAL / 物理地址）。
 * 分工声明 (Scope)      : 与 `FC_DL_TableLookupDescending` 分工：区间定位归那件、
 *                         最近点归本件；与 `FC_DL_TableIndexBinarySearch` 分工：
 *                         二分只适用于有序大表，本件为无序/小表通用件。
 * 来源标签 (Source Tag) : 原创实现（无外部代码引入）
 * 码表     (Codes)      : 本件不占用全局数字码位；出口为 BOOL + INT + LREAL +
 *                         本文件内定义 enum E_DL_TblNearErr（全库唯一）。
 * 红线自检 (Redline)    : R1 ✓ 零 GVL/VAR_EXTERNAL ｜ R2 ✓ 零 %I/%Q/%M ｜ R3 ✓ 纯 IEC 61131-3
 *                         R4 ✓ 点数域闸 + 全表非有限双判 + 距离非负复检 ｜ R5 ✓ 声明逐行同行双语注释
 *                         R6 N/A（纯函数无状态机） ｜ R7 N/A（无实例调用）
 * 修订历史 (Revision)   : 2026-11-23  v1.0.0  R77 首版（批次 B3 · 序号 2）
 * 验收向量 (Acceptance) : ① afX=[10,20,30], iCount=3, fXin=23.0 → iIndex=2, fDist=3.0, eOk, TRUE；
 *                         ② afX=[10,20,30], fXin=25.0 → 与 20/30 等距 5.0 → iIndex=2（取较小下标）, fDist=5.0；
 *                         ③ afX=[10,20,30], fXin=100.0 → iIndex=3, fDist=70.0；
 *                         ④ iCount=0 → 返回 FALSE, iIndex=0, eBadCount；
 *                         ⑤ afX[2]=NaN → 返回 FALSE, eNonFinite。
 *==============================================================================*)

(*-----------------------------------------------------------------------------
 * 枚举: E_DL_TblNearErr（最近节点查找错误码，归属 DL_MathData，与本件同文件，全库唯一属主）
 *----------------------------------------------------------------------------*)
TYPE E_DL_TblNearErr :
(
    eOk        := 0,   // 信息级：查找完成 / Info: lookup completed
    eBadCount  := 1,   // 故障级：点数越域 / Fault: point count out of domain
    eNonFinite := 2    // 故障级：查询点或表元素非有限 / Fault: query or table entry non-finite
);
END_TYPE

FUNCTION FC_DL_TableLookupNearestIndex : BOOL
VAR_INPUT
    afX    : ARRAY[1..32] OF LREAL;  // 节点表（无需有序） [任意工程量] / Node table, order not required
    iCount : INT;                    // 有效点数（1..32） [个] / Valid point count, 1..32
    fXin   : LREAL;                  // 查询点 [同 afX 单位] / Query value, same unit as afX
END_VAR
VAR_OUTPUT
    iIndex   : INT;    // 最近节点下标（1..iCount） [-] / Nearest node index
    fDist    : LREAL;  // 最小绝对距离 [同 afX 单位] / Minimum absolute distance
    eErrCode : E_DL_TblNearErr; // 错误码出口 [-] / Error code outlet
END_VAR
VAR
    _i       : INT;    // 循环下标 [-] / Loop index
    _iBest   : INT;    // 当前最优下标 [-] / Current best index
    _bNonFin : BOOL;   // 非有限标志 [-] / Non-finite flag
    _fBest   : LREAL;  // 当前最优距离 [同 afX 单位] / Current best distance
    _fCur    : LREAL;  // 当前候选距离 [同 afX 单位] / Current candidate distance
END_VAR
VAR CONSTANT
    DL_TNC_CNT_MIN : INT := 1;        // 点数下限 [个] / Count lower bound
    DL_TNC_CNT_MAX : INT := 32;       // 点数上限（数组容量） [个] / Count upper bound
    DL_TNC_ZERO    : LREAL := 0.0;    // 零与距离下限 [-] / Zero and distance lower bound
    DL_TNC_BIG     : LREAL := 1.0E30; // 初值大数（保证首次必被更替） [-] / Large seed ensuring first replacement
END_VAR

(* —— 段 0：出口预置安全值 —— *)
FC_DL_TableLookupNearestIndex := FALSE;            // 返回值预置无效 / Return preset invalid
iIndex   := 0;                                     // 下标哨兵 0 / Index sentinel
fDist    := DL_TNC_ZERO;                           // 距离哨兵 0 / Distance sentinel
eErrCode := E_DL_TblNearErr.eBadCount;             // 预置最严码 / Preset strictest code

(* —— 段 1：点数域闸 —— *)
IF (iCount < DL_TNC_CNT_MIN) OR (iCount > DL_TNC_CNT_MAX) THEN
    RETURN;                                        // 点数越域：保持故障码与哨兵 / Count out of domain
END_IF

(* —— 段 2：非有限域闸（查询点 + 全部表元素逐项枚举） —— *)
_bNonFin := (fXin <> fXin) OR ((fXin - fXin) <> DL_TNC_ZERO);   // 查询点非有限 / Query non-finite
_i := 1;
WHILE _i <= iCount DO
    IF (afX[_i] <> afX[_i]) OR ((afX[_i] - afX[_i]) <> DL_TNC_ZERO) THEN
        _bNonFin := TRUE;                          // 表元素非有限 / Table entry non-finite
    END_IF
    _i := _i + 1;
END_WHILE
IF _bNonFin THEN
    eErrCode := E_DL_TblNearErr.eNonFinite;        // 故障级码 / Fault-level code
    RETURN;
END_IF

(* —— 段 3：最小绝对距离扫描（严格 < 比较 → 并列时保留较小下标） —— *)
_iBest := 1;                                       // 最优下标初值 / Best index seed
_fBest := DL_TNC_BIG;                              // 最优距离初值 / Best distance seed
_i     := 1;
WHILE _i <= iCount DO
    _fCur := ABS(afX[_i] - fXin);                  // 绝对距离（非负） / Absolute distance
    IF _fCur < _fBest THEN
        _fBest := _fCur;                           // 更优距离 / Better distance
        _iBest := _i;                              // 更新下标 / Update index
    END_IF
    _i := _i + 1;
END_WHILE

(* —— 段 4：结果复检（下标域 + 距离非负且有限） —— *)
IF (_iBest < DL_TNC_CNT_MIN) OR (_iBest > iCount) THEN
    eErrCode := E_DL_TblNearErr.eBadCount;         // 下标越域：内部不一致 / Index out of domain
    RETURN;
END_IF
IF (_fBest <> _fBest) OR ((_fBest - _fBest) <> DL_TNC_ZERO) OR (_fBest < DL_TNC_ZERO) THEN
    eErrCode := E_DL_TblNearErr.eNonFinite;        // 距离异常 / Abnormal distance
    RETURN;
END_IF

iIndex   := _iBest;                                // 导出最近下标 / Export nearest index
fDist    := _fBest;                                // 导出最小距离 / Export minimum distance
eErrCode := E_DL_TblNearErr.eOk;                   // 信息级成功 / Info success
FC_DL_TableLookupNearestIndex := TRUE;             // 查找可信 / Lookup trustworthy

END_FUNCTION

(* ---- FC_DL_TableReverseLookupX.st ---- *)
(*==============================================================================
 * 组件名称 (Component)  : FC_DL_TableReverseLookupX
 * 所属子库 (Sublibrary) : DL_MathData
 * 当前版本 (Version)    : 1.0.0
 * 兼容性   (Platform)   : CODESYS 3.5+ / TwinCAT 3 / 汇川 InoProShop / 施耐德 Machine Expert
 *                         仅依赖 IEC 61131-3 标准数学（ABS / MIN / MAX），零厂商私有库
 * 功能描述 (Function)   : 由 Y 反查 X（单调表反解）。给定单调的 afY 表与对应 afX 表，
 *                         输入 fYin 反求 X：
 *                           ① 先做**全表单调性校验**：逐对比较相邻 afY，全升或全降才合法；
 *                             平坦段（|ΔY| < 1E-9）允许多个连续，但整表必须同向；
 *                           ② 再在 afY 中定位区间并按线性插值反解 X：
 *                              x = x_i + (x_{i+1} - x_i) × (yin - y_i) / (y_{i+1} - y_i)
 *                           ③ fYin 超出 afY 范围 → 钳到端点并置 bClamped（不外推，
 *                             反解外推在工艺上几乎总是错的）。
 *                         用途：由实测压力反查饱和温度、由输出反馈反查指令给定（阀位反解）。
 * 接口     (Interface)  : 输入 afY 单调表 [Y 单位]、afX 对应表 [X 单位]、
 *                         iCount 有效点数 [个]（2..32）、fYin 查询值 [Y 单位]；
 *                         输出 fXout 反解结果 [X 单位]、iSeg 区间下标、
 *                         bIncreasing 表是否升序（诊断）、bClamped 越界钳位回执、
 *                         eErrCode（E_DL_TblRevErr）；
 *                         返回值 = bValid 反解可信标志（TRUE = fXout 可信）。
 * 边界     (Boundary)   : ① 属主边界：只做单调表反解，不做非单调表的「多值择一」
 *                         （非单调 → 故障级 eNotMonotonic，**拒绝而非猜测**）。
 *                         ② 点数域闸 2..32；越域 → 故障级 eBadCount。
 *                         ③ 非有限双判：查询值 + afY 与 afX 双表全部元素逐项枚举。
 *                         ④ 段宽（ΔY）近似零 → 该段内反解取左端 X 并置信息级 eDegenerateSeg
 *                         （除零防护；平坦段反解本身欠定，取左端是确定性选择）。
 *                         ⑤ 单调性校验含符号一致性：先用首对非平坦段定方向，
 *                         后续任何反向段即判 eNotMonotonic。
 *                         ⑥ 零全局耦合（无 GVL / VAR_EXTERNAL / 物理地址）。
 * 分工声明 (Scope)      : 与 `FC_DL_TableIndexBinarySearch` 分工：正查（X→区间）归那件、
 *                         反查（Y→X）归本件；与 `FC_DL_InterpHoldLast` 分工：
 *                         保持型正查归那件，本件同样禁止外推。
 * 来源标签 (Source Tag) : 原创实现（无外部代码引入）
 * 码表     (Codes)      : 本件不占用全局数字码位；出口为 BOOL + LREAL + INT + 2×BOOL +
 *                         本文件内定义 enum E_DL_TblRevErr（全库唯一）。
 * 红线自检 (Redline)    : R1 ✓ 零 GVL/VAR_EXTERNAL ｜ R2 ✓ 零 %I/%Q/%M ｜ R3 ✓ 纯 IEC 61131-3
 *                         R4 ✓ 双表全元素非有限双判 + ΔY 判零（除零防护）+ 单调性校验 + 越界钳位 ｜ R5 ✓ 声明逐行同行双语注释
 *                         R6 N/A（纯函数无状态机） ｜ R7 N/A（无实例调用）
 * 修订历史 (Revision)   : 2026-11-23  v1.0.0  R77 首版（批次 B3 · 序号 7）
 * 验收向量 (Acceptance) : ① afY=[0,100,200], afX=[0,10,20], iCount=3, fYin=150 →
 *                         bIncreasing=TRUE, iSeg=2, fXout=15.0（容差 1E-9）, eOk, TRUE；
 *                         ② afY=[200,100,0]（降序）, afX=[0,10,20], fYin=150 →
 *                         bIncreasing=FALSE, fXout=5.0（容差 1E-9）；
 *                         ③ afY=[0,100,200], fYin=999 → fXout=20.0（钳到末端点）, bClamped=TRUE；
 *                         ④ afY=[0,100,50]（非单调）→ 返回 FALSE, eNotMonotonic；
 *                         ⑤ fYin=NaN → 返回 FALSE, eNonFinite。
 *==============================================================================*)

(*-----------------------------------------------------------------------------
 * 枚举: E_DL_TblRevErr（单调表反解错误码，归属 DL_MathData，与本件同文件，全库唯一属主）
 *----------------------------------------------------------------------------*)
TYPE E_DL_TblRevErr :
(
    eOk            := 0,   // 信息级：反解完成 / Info: reverse lookup done
    eDegenerateSeg := 1,   // 信息级：ΔY 近似零，取左端 X / Info: flat segment, left X used
    eBadCount      := 2,   // 故障级：点数越域 / Fault: point count out of domain
    eNonFinite     := 3,   // 故障级：任一入参或表元素非有限 / Fault: any input or table entry non-finite
    eNotMonotonic  := 4    // 故障级：表非单调，反解多值 / Fault: non-monotonic table, multiple solutions
);
END_TYPE

FUNCTION FC_DL_TableReverseLookupX : BOOL
VAR_INPUT
    afY    : ARRAY[1..32] OF LREAL;  // 单调值表 [Y 单位] / Monotonic value table in Y
    afX    : ARRAY[1..32] OF LREAL;  // 对应自变量表 [X 单位] / Corresponding argument table in X
    iCount : INT;                    // 有效点数（2..32） [个] / Valid point count, 2..32
    fYin   : LREAL;                  // 查询值 [Y 单位] / Query value in Y
END_VAR
VAR_OUTPUT
    fXout       : LREAL;  // 反解结果 [X 单位] / Reverse-solved X
    iSeg        : INT;    // 区间下标（1..iCount-1） [-] / Segment index
    bIncreasing : BOOL;   // 表是否升序（诊断） [-] / Whether the table is ascending
    bClamped    : BOOL;   // 越界钳位回执 [-] / Out-of-range clamp receipt
    eErrCode    : E_DL_TblRevErr; // 错误码出口 [-] / Error code outlet
END_VAR
VAR
    _i        : INT;    // 循环下标 [-] / Loop index
    _iSeg     : INT;    // 命中区间下标 [-] / Hit segment index
    _bFound   : BOOL;   // 区间命中标志 [-] / Segment found flag
    _bNonFin  : BOOL;   // 非有限标志 [-] / Non-finite flag
    _bInc     : BOOL;   // 方向已定标志 [-] / Direction determined flag
    _bUp      : BOOL;   // 方向：升序 = TRUE [-] / Direction, ascending equals TRUE
    _fDy      : LREAL;  // ΔY（分母） [Y 单位] / Delta Y denominator
    _fRatio   : LREAL;  // 段内比例 [-] / In-segment ratio
END_VAR
VAR CONSTANT
    DL_TRC_CNT_MIN : INT := 2;        // 点数下限 [个] / Count lower bound
    DL_TRC_CNT_MAX : INT := 32;       // 点数上限（数组容量） [个] / Count upper bound
    DL_TRC_TINY    : LREAL := 1.0E-9; // ΔY 近似零阈值（平坦段） [Y 单位] / Flat segment threshold
    DL_TRC_ZERO    : LREAL := 0.0;    // 零基准与比例下限 [-] / Zero base and ratio lower bound
    DL_TRC_ONE     : LREAL := 1.0;    // 比例上限 [-] / Ratio upper bound
END_VAR

(* —— 段 0：出口预置安全值 —— *)
FC_DL_TableReverseLookupX := FALSE;                // 返回值预置无效 / Return preset invalid
fXout       := DL_TRC_ZERO;                        // 结果哨兵 0 / Result sentinel
iSeg        := 0;                                  // 下标哨兵 / Index sentinel
bIncreasing := FALSE;                              // 方向标志预置否 / Direction preset false
bClamped    := FALSE;                              // 钳位回执预置否 / Clamp receipt preset false
eErrCode    := E_DL_TblRevErr.eBadCount;           // 预置最严码 / Preset strictest code

(* —— 段 1：点数域闸 —— *)
IF (iCount < DL_TRC_CNT_MIN) OR (iCount > DL_TRC_CNT_MAX) THEN
    RETURN;
END_IF

(* —— 段 2：非有限域闸（查询值 + afY 与 afX 双表逐项枚举） —— *)
_bNonFin := (fYin <> fYin) OR ((fYin - fYin) <> DL_TRC_ZERO);
_i := 1;
WHILE _i <= iCount DO
    IF (afY[_i] <> afY[_i]) OR ((afY[_i] - afY[_i]) <> DL_TRC_ZERO) THEN
        _bNonFin := TRUE;                          // Y 表元素非有限 / Y entry non-finite
    END_IF
    IF (afX[_i] <> afX[_i]) OR ((afX[_i] - afX[_i]) <> DL_TRC_ZERO) THEN
        _bNonFin := TRUE;                          // X 表元素非有限 / X entry non-finite
    END_IF
    _i := _i + 1;
END_WHILE
IF _bNonFin THEN
    eErrCode := E_DL_TblRevErr.eNonFinite;
    RETURN;
END_IF

(* —— 段 3：全表单调性校验（首对非平坦段定向，后续任一反向即判非单调） —— *)
_bInc   := FALSE;                                  // 方向尚未确定 / Direction not yet determined
_bUp    := TRUE;                                   // 方向暂定升序 / Direction provisionally ascending
_i      := 1;
WHILE _i < iCount DO
    _fDy := afY[_i + 1] - afY[_i];                 // 相邻差 / Adjacent difference
    IF ABS(_fDy) >= DL_TRC_TINY THEN
        IF NOT _bInc THEN
            _bInc := TRUE;                         // 首对非平坦段定方向 / First non-flat pair determines direction
            _bUp  := (_fDy > DL_TRC_ZERO);
        ELSE
            IF (_bUp AND (_fDy < DL_TRC_ZERO)) OR ((NOT _bUp) AND (_fDy > DL_TRC_ZERO)) THEN
                eErrCode := E_DL_TblRevErr.eNotMonotonic;   // 方向反转：非单调 / Direction reversal
                RETURN;
            END_IF
        END_IF
    END_IF
    _i := _i + 1;
END_WHILE
IF NOT _bInc THEN
    eErrCode := E_DL_TblRevErr.eNotMonotonic;      // 全表平坦：反解多值 / Fully flat: multiple solutions
    RETURN;
END_IF
bIncreasing := _bUp;                               // 导出方向诊断 / Export direction diagnostic

(* —— 段 4：越界钳位（低于首端 / 高于末端，均不外推） —— *)
IF _bUp THEN
    IF fYin <= afY[1] THEN
        fXout    := afX[1];
        iSeg     := 1;
        bClamped := TRUE;
        eErrCode := E_DL_TblRevErr.eOk;
        FC_DL_TableReverseLookupX := TRUE;
        RETURN;
    END_IF
    IF fYin >= afY[iCount] THEN
        fXout    := afX[iCount];
        iSeg     := iCount - 1;
        bClamped := TRUE;
        eErrCode := E_DL_TblRevErr.eOk;
        FC_DL_TableReverseLookupX := TRUE;
        RETURN;
    END_IF
ELSE
    IF fYin >= afY[1] THEN
        fXout    := afX[1];
        iSeg     := 1;
        bClamped := TRUE;
        eErrCode := E_DL_TblRevErr.eOk;
        FC_DL_TableReverseLookupX := TRUE;
        RETURN;
    END_IF
    IF fYin <= afY[iCount] THEN
        fXout    := afX[iCount];
        iSeg     := iCount - 1;
        bClamped := TRUE;
        eErrCode := E_DL_TblRevErr.eOk;
        FC_DL_TableReverseLookupX := TRUE;
        RETURN;
    END_IF
END_IF

(* —— 段 5：区间定位（按方向取包围区间） —— *)
_i      := 1;
_bFound := FALSE;
_iSeg   := 1;
WHILE (_i < iCount) AND (NOT _bFound) DO
    IF _bUp THEN
        IF (fYin >= afY[_i]) AND (fYin <= afY[_i + 1]) THEN
            _bFound := TRUE;
            _iSeg   := _i;
        END_IF
    ELSE
        IF (fYin <= afY[_i]) AND (fYin >= afY[_i + 1]) THEN
            _bFound := TRUE;
            _iSeg   := _i;
        END_IF
    END_IF
    IF NOT _bFound THEN
        _i := _i + 1;
    END_IF
END_WHILE
IF NOT _bFound THEN
    eErrCode := E_DL_TblRevErr.eNotMonotonic;      // 未命中：与单调性矛盾 / Not found: contradicts monotonicity
    RETURN;
END_IF

(* —— 段 6：ΔY 判零后反解（除零防护） —— *)
_fDy := afY[_iSeg + 1] - afY[_iSeg];               // ΔY / Delta Y
IF ABS(_fDy) < DL_TRC_TINY THEN
    fXout    := afX[_iSeg];                        // 平坦段：取左端 X（确定性选择） / Flat: deterministic left X
    eErrCode := E_DL_TblRevErr.eDegenerateSeg;     // 信息级码 / Info code
ELSE
    _fRatio  := (fYin - afY[_iSeg]) / _fDy;        // 段内比例 / In-segment ratio
    _fRatio  := MIN(MAX(_fRatio, DL_TRC_ZERO), DL_TRC_ONE);   // 显式约束 0..1 / Constrain 0..1
    fXout    := afX[_iSeg] + (afX[_iSeg + 1] - afX[_iSeg]) * _fRatio;   // 线性反解 X / Linear reverse solve
    eErrCode := E_DL_TblRevErr.eOk;                // 信息级成功 / Info success
END_IF
iSeg := _iSeg;

(* —— 段 7：结果非有限复检兜底 —— *)
IF (fXout <> fXout) OR ((fXout - fXout) <> DL_TRC_ZERO) THEN
    fXout    := DL_TRC_ZERO;
    iSeg     := 0;
    eErrCode := E_DL_TblRevErr.eNonFinite;
    RETURN;
END_IF

FC_DL_TableReverseLookupX := TRUE;                 // 反解有效 / Reverse lookup valid

END_FUNCTION

(* ---- FC_DL_ThermocoupleLinearization.st ---- *)
(*
  ==================================================================
  组件名 Component  : FC_DL_ThermocoupleLinearization
  分类   Category   : DL_MathData
  复杂度 Complexity  : 中
  版本   Version    : 1.0.0
  功能   Purpose    : 热电偶 mV↔温度双向线性化（K / N / S 三型）。内部按公开
                      ITS-90 参考分度表特征点（100 摄氏度步距锚点）做折线
                      插值，正向（温度→mV）与反向（mV→温度）共用同一单调
                      锚点表，域外钳位并置信息级，未知型别 / 非法方向 / 表
                      单调破坏判故障级。与 RtdLinearization / TempUnitConvert
                      / NtcTempScan 三分工边界按 ROADMAP 1083 行写死。
  来源   Source     : roadmap-p1（R56 评估项落地）
  溯源   Origin     : 锚点数值取自公开 ITS-90 热电偶参考分度表（clean-room
                      整理），插值算法为自研折线实现，未复制 NIST 数据库
                      程序或任何厂商私有库源码。
  精度声明 Precision : 100 摄氏度步距折线插值，K / N 型 0..1000 摄氏度段典型
                      误差 ±1.5 K 量级（S 型低温段略宽）；非 NIST 全阶多项式
                      ——全阶系数升级挂编译验证债（入库后另行立项复核）。
  平台   Platform   : 纯 IEC 61131-3，CODESYS / TwinCAT / InoProShop 通用
  分工声明 Split     : 与 FC_DL_RtdLinearization 分工——Rtd 为铂电阻 Callendar-
                      Van Dusen 方程口径；与 FC_DL_TempUnitConvert 分工——
                      后者只做摄氏 / 华氏 / 开尔文单位换算；与 FB_DL_NtcTempScan
                      分工——Ntc 为 NTC 热敏电阻扫描查表；本件只做热电偶
                      mV↔温度双向线性化。
  作者   Author     : 道莅代码库 · PLC 编程专家（R58）
  ------------------------------------------------------------------
  功能说明  : 输入 fIn 按方向解释：eTempToMv 时 fIn 为摄氏度 [摄氏度]，返回
              毫伏 [毫伏]；eMvToTemp 时 fIn 为毫伏 [毫伏]，返回摄氏度 [摄氏度]。
              域闸门四段式（R45）：预置 → 非有限 / 型别 / 方向 / 单调性闸 →
              域内插值 → 结果非有限复检兜底。
  输出约定  : bError = TRUE 仅故障级（非有限 / 型别非法 / 方向非法 / 表单调
              破坏）；bClamped = TRUE 为信息级域外钳位（不置 bError），此时
              返回值为钳位端点值。
  修订记录  : 2026-11-21 v1.0.0 首次入库（R58 批 1 · 序号 3）
*)

(*-----------------------------------------------------------------------------
 * 枚举: E_DL_TcKind（唯一属主 = 本文件，R67 全库唯一断言）
 * 含义: 支持的热电偶型别。
 *----------------------------------------------------------------------------*)
TYPE E_DL_TcKind :
(
    eTcK := 0, // K 型热电偶（镍铬 - 镍硅）/ the type K thermocouple
    eTcN := 1, // N 型热电偶（镍铬硅 - 镍硅）/ the type N thermocouple
    eTcS := 2  // S 型热电偶（铂铑 10 - 铂）/ the type S thermocouple
);
END_TYPE

(*-----------------------------------------------------------------------------
 * 枚举: E_DL_TcDir（唯一属主 = 本文件，R67 全库唯一断言）
 * 含义: 线性化方向。
 *----------------------------------------------------------------------------*)
TYPE E_DL_TcDir :
(
    eTempToMv := 0, // 正向：温度 → 毫伏 / the forward direction, temperature to millivolt
    eMvToTemp := 1  // 反向：毫伏 → 温度 / the reverse direction, millivolt to temperature
);
END_TYPE

(*-----------------------------------------------------------------------------
 * 枚举: E_DL_TlcCause（唯一属主 = 本文件，R67 全库唯一断言；零码位范式，
 *       收口派号前不写 16# 事件码，故障出口 = BOOL + ENUM）
 * 含义: 线性化结果成因（1..3 故障级 / 4 信息级）。
 *----------------------------------------------------------------------------*)
TYPE E_DL_TlcCause :
(
    eTlcNone         := 0, // 无成因 / no cause
    eTlcNonFinite    := 1, // 输入或结果非有限（故障级，与 bError 配对）/ a non finite input or result
    eTlcKindBad      := 2, // 型别非法或锚点表单调破坏（故障级，与 bError 配对）/ an unknown kind or a monotony break
    eTlcDirBad       := 3, // 方向非法（故障级，与 bError 配对）/ an illegal direction
    eTlcRangeClamped := 4  // 域外钳位（信息级，不置 bError）/ an out of range clamp, informational
);
END_TYPE

FUNCTION FC_DL_ThermocoupleLinearization : LREAL
VAR_INPUT
    fIn  : LREAL; // 输入量：正向为摄氏度 [摄氏度]，反向为毫伏 [毫伏] / the input, temperature in celsius forward or millivolt reverse
    eKind: E_DL_TcKind; // 热电偶型别选择 [枚举] / the thermocouple kind selector
    eDir : E_DL_TcDir;  // 线性化方向选择 [枚举] / the linearization direction selector
END_VAR
VAR_OUTPUT
    bError   : BOOL; // 故障标志，仅故障级置位 / the fault flag, fault grade only
    bClamped : BOOL; // 域外钳位发生（信息级，不置 bError）[-] / an out of range clamp happened, informational
    eCause   : E_DL_TlcCause; // 成因出口 [枚举] / the cause outlet
END_VAR
VAR
    afT    : ARRAY[0..17] OF LREAL; // 工作锚点温度表 [摄氏度] / the working anchor temperature table [degree celsius]
    afM    : ARRAY[0..17] OF LREAL; // 工作锚点热电势表 [毫伏] / the working anchor millivolt table [millivolt]
    nAnch  : DINT;  // 工作表有效锚点数 [个] / the valid anchor count of the working table
    nI     : DINT;  // 锚点遍历索引 [个] / the anchor loop index
    nSeg   : DINT;  // 命中段索引 [段] / the hit segment index
    lrX    : LREAL; // 工作量（已判向后的输入）[混合] / the working value after the direction verdict
    lrDen  : LREAL; // 命中段分母（锚点差）[混合] / the hit segment denominator
    lrRes  : LREAL; // 结果工作量 [混合] / the result working value
    bBad   : BOOL;  // 故障级闸命中工作量 [-] / the fault gate hit work flag
END_VAR
VAR CONSTANT
    aTkT : ARRAY[0..14] OF LREAL := [-100.0, 0.0, 100.0, 200.0, 300.0, 400.0, 500.0, 600.0, 700.0, 800.0, 900.0, 1000.0, 1100.0, 1200.0, 1300.0]; // K 型锚点温度表 [摄氏度]，严格递增 / the type K anchor temperatures, strictly increasing
    aTkM : ARRAY[0..14] OF LREAL := [-3.554, 0.0, 4.096, 8.138, 12.209, 16.397, 20.644, 24.905, 29.129, 33.275, 37.326, 41.276, 45.119, 48.838, 52.398]; // K 型锚点热电势表 [毫伏]，严格递增 / the type K anchor millivolts, strictly increasing
    aTnT : ARRAY[0..14] OF LREAL := [-100.0, 0.0, 100.0, 200.0, 300.0, 400.0, 500.0, 600.0, 700.0, 800.0, 900.0, 1000.0, 1100.0, 1200.0, 1300.0]; // N 型锚点温度表 [摄氏度]，严格递增 / the type N anchor temperatures, strictly increasing
    aTnM : ARRAY[0..14] OF LREAL := [-2.655, 0.0, 2.774, 5.913, 9.341, 12.974, 16.748, 20.644, 24.639, 28.608, 32.542, 36.382, 40.103, 43.770, 47.348]; // N 型锚点热电势表 [毫伏]，严格递增 / the type N anchor millivolts, strictly increasing
    aTsT : ARRAY[0..17] OF LREAL := [0.0, 100.0, 200.0, 300.0, 400.0, 500.0, 600.0, 700.0, 800.0, 900.0, 1000.0, 1100.0, 1200.0, 1300.0, 1400.0, 1500.0, 1600.0, 1700.0]; // S 型锚点温度表 [摄氏度]，严格递增 / the type S anchor temperatures, strictly increasing
    aTsM : ARRAY[0..17] OF LREAL := [0.0, 0.646, 1.441, 2.323, 3.259, 4.233, 5.239, 6.274, 7.345, 8.448, 9.587, 10.754, 11.947, 13.159, 14.373, 15.582, 16.777, 17.942]; // S 型锚点热电势表 [毫伏]，严格递增 / the type S anchor millivolts, strictly increasing
END_VAR

// 段 1｜返回值与错误状态预置安全值（四段式第一段，R45）/ segment 1, preset the return and error states
FC_DL_ThermocoupleLinearization := 0.0; // 返回值预置 0.0 / preset the return to the safe zero
bError   := FALSE; // 故障标志预置假 / preset the fault flag false
bClamped := FALSE; // 钳位标志预置假 / preset the clamp flag false
eCause   := E_DL_TlcCause.eTlcNone; // 成因预置无 / preset the cause none
bBad     := FALSE; // 故障闸工作量预置假 / preset the fault work flag false

// 段 2｜非有限拦截（自反双判据，R79）/ segment 2, the non finite interception
IF (fIn <> fIn) OR ((fIn - fIn) <> (fIn - fIn)) THEN // 输入非有限 / a non finite input
    bBad   := TRUE; // 置故障闸 / raise the fault gate
    eCause := E_DL_TlcCause.eTlcNonFinite; // 故障级成因（R45 配对）/ the fault cause
END_IF

// 段 3｜型别装表 + 方向闸 + 表单调自检 / segment 3, the table loading, the direction gate and the monotony self check
IF NOT bBad THEN // 非有限未命中才装表 / load the table only when finite
    CASE eKind OF // 按型别装工作表（其余锚点槽保持缺省零，不在有效域内使用）/ load the working table by kind
    E_DL_TcKind.eTcK: // K 型 / the type K
        nAnch := 15; // 有效锚点数 / the valid anchor count
        FOR nI := 0 TO 14 DO // 固定界复制 / the fixed bound copy
            afT[nI] := aTkT[nI]; // 装温度锚点 / load the temperature anchor
            afM[nI] := aTkM[nI]; // 装热电势锚点 / load the millivolt anchor
        END_FOR
    E_DL_TcKind.eTcN: // N 型 / the type N
        nAnch := 15; // 有效锚点数 / the valid anchor count
        FOR nI := 0 TO 14 DO // 固定界复制 / the fixed bound copy
            afT[nI] := aTnT[nI]; // 装温度锚点 / load the temperature anchor
            afM[nI] := aTnM[nI]; // 装热电势锚点 / load the millivolt anchor
        END_FOR
    E_DL_TcKind.eTcS: // S 型 / the type S
        nAnch := 18; // 有效锚点数 / the valid anchor count
        FOR nI := 0 TO 17 DO // 固定界复制 / the fixed bound copy
            afT[nI] := aTsT[nI]; // 装温度锚点 / load the temperature anchor
            afM[nI] := aTsM[nI]; // 装热电势锚点 / load the millivolt anchor
        END_FOR
    ELSE // 未知型别兜底（R128）/ the unknown kind fallback
        nAnch  := 0; // 不装表 / no table
        bBad   := TRUE; // 置故障闸 / raise the fault gate
        eCause := E_DL_TlcCause.eTlcKindBad; // 故障级成因 / the fault cause
    END_CASE
    IF (NOT bBad) AND (nAnch >= 2) THEN // 表已装且至少两锚点才自检 / self check with a loaded table
        FOR nI := 0 TO nAnch - 2 DO // 逐段单调自检（防御深，常量表本应单调）/ the per segment monotony self check, defense in depth
            IF (afT[nI + 1] <= afT[nI]) OR (afM[nI + 1] <= afM[nI]) THEN // 单调破坏 / a monotony break
                bBad   := TRUE; // 置故障闸 / raise the fault gate
                eCause := E_DL_TlcCause.eTlcKindBad; // 故障级成因（表损坏归型别成因）/ the fault cause, a broken table maps to the kind cause
            END_IF
        END_FOR
    END_IF
END_IF

// 段 4｜方向闸与双向插值（域外钳位信息级，除子单调已证大于零）/ segment 4, the direction gate and the bidirectional interpolation
IF NOT bBad THEN // 无故障才插值 / interpolate only without a fault
    CASE eDir OF // 方向闸（含非法方向兜底 R128）/ the direction gate with the illegal fallback
    E_DL_TcDir.eTempToMv: // 正向：温度→毫伏 / the forward direction
        lrX := fIn; // 工作量为摄氏度 / the working value in celsius
        IF lrX < afT[0] THEN // 低于域下界 / below the floor
            lrX := afT[0]; // 钳到下端点 / clamp to the lower anchor
            bClamped := TRUE; // 信息级钳位 / the informational clamp
        ELSIF lrX > afT[nAnch - 1] THEN // 高于域上界 / above the bound
            lrX := afT[nAnch - 1]; // 钳到上端点 / clamp to the upper anchor
            bClamped := TRUE; // 信息级钳位 / the informational clamp
        END_IF
        nSeg := nAnch - 2; // 段索引预置末段（上端点命中）/ preset the last segment
        FOR nI := 0 TO nAnch - 2 DO // 有界段搜索（命中即出，无死循环）/ the bounded segment search
            IF lrX <= afT[nI + 1] THEN // 命中段 / a hit segment
                nSeg := nI; // 记段索引 / record the segment
                EXIT; // 提前出循环 / leave early
            END_IF
        END_FOR
        lrDen := afT[nSeg + 1] - afT[nSeg]; // 温差分母 [摄氏度] / the temperature denominator
        IF lrDen > 1.0E-12 THEN // 除子护栏（单调自检已证，防御深）/ the divisor guard
            lrRes := afM[nSeg] + (lrX - afT[nSeg]) * (afM[nSeg + 1] - afM[nSeg]) / lrDen; // 折线插值 / the linear interpolation
        ELSE // 分母退化（不可达路径兜底）/ the degenerate divisor, unreachable
            bBad   := TRUE; // 置故障闸 / raise the fault gate
            eCause := E_DL_TlcCause.eTlcKindBad; // 故障级成因 / the fault cause
        END_IF
    E_DL_TcDir.eMvToTemp: // 反向：毫伏→温度 / the reverse direction
        lrX := fIn; // 工作量为毫伏 / the working value in millivolt
        IF lrX < afM[0] THEN // 低于域下界 / below the floor
            lrX := afM[0]; // 钳到下端点 / clamp to the lower anchor
            bClamped := TRUE; // 信息级钳位 / the informational clamp
        ELSIF lrX > afM[nAnch - 1] THEN // 高于域上界 / above the bound
            lrX := afM[nAnch - 1]; // 钳到上端点 / clamp to the upper anchor
            bClamped := TRUE; // 信息级钳位 / the informational clamp
        END_IF
        nSeg := nAnch - 2; // 段索引预置末段 / preset the last segment
        FOR nI := 0 TO nAnch - 2 DO // 有界段搜索 / the bounded segment search
            IF lrX <= afM[nI + 1] THEN // 命中段 / a hit segment
                nSeg := nI; // 记段索引 / record the segment
                EXIT; // 提前出循环 / leave early
            END_IF
        END_FOR
        lrDen := afM[nSeg + 1] - afM[nSeg]; // 热电势差分母 [毫伏] / the millivolt denominator
        IF lrDen > 1.0E-12 THEN // 除子护栏（单调自检已证，防御深）/ the divisor guard
            lrRes := afT[nSeg] + (lrX - afM[nSeg]) * (afT[nSeg + 1] - afT[nSeg]) / lrDen; // 反向折线插值 / the reverse interpolation
        ELSE // 分母退化（不可达路径兜底）/ the degenerate divisor, unreachable
            bBad   := TRUE; // 置故障闸 / raise the fault gate
            eCause := E_DL_TlcCause.eTlcKindBad; // 故障级成因 / the fault cause
        END_IF
    ELSE // 非法方向兜底（R128）/ the illegal direction fallback
        bBad   := TRUE; // 置故障闸 / raise the fault gate
        eCause := E_DL_TlcCause.eTlcDirBad; // 故障级成因 / the fault cause
    END_CASE
END_IF

// 段 5｜结果非有限复检兜底（防御纵深，正常路径不可达）/ segment 5, the result recheck as defense in depth
IF (NOT bBad) AND ((lrRes <> lrRes) OR ((lrRes - lrRes) <> (lrRes - lrRes))) THEN // 结果非有限 / a non finite result
    bBad   := TRUE; // 置故障闸 / raise the fault gate
    eCause := E_DL_TlcCause.eTlcNonFinite; // 故障级成因 / the fault cause
END_IF
IF bBad THEN // 故障出口 / the fault outlet
    FC_DL_ThermocoupleLinearization := 0.0; // 返回预置安全值 / return the safe zero
    bError := TRUE; // 置故障标志（R45 配对）/ raise the fault flag
ELSE // 正常出口 / the normal outlet
    FC_DL_ThermocoupleLinearization := lrRes; // 返回插值结果 / return the interpolation result
END_IF
END_FUNCTION

(* ---- FC_DL_TimeUnitConvert.st ---- *)
(*==============================================================================
 * 组件名称 : FC_DL_TimeUnitConvert ｜ 子库 : DL_MathData ｜ v1.0.0 ｜ 2026-11-23
 * 平台     : CODESYS 3.5 / TwinCAT 3 / InoProShop / Machine Expert（纯 IEC，无厂商库）
 * 功能简介 : 时间单位 s / min / h 两两互转。源/目标由枚举对单向选择，
 *            单向基准链（先归一到 s）使公式域固定为 3+3 条分支。
 * 契约     : 返回换算结果 [目标单位]；枚举非法（越界值）返回 0.0；
 *            除数为编译期非零常量，无除零风险；纯函数无状态。
 * 依赖     : 无 DL_ 内部依赖（本批自足实现）
 * 红线自检 : R1 零全局 R2 零%I/%Q R3 纯IEC R4 枚举越界拒收返 0 + 常量除数
 *            R5 全变量与枚举项双语同行注释 R6 N/A（无状态机） R7 N/A
 * 修订历史 : 2026-11-23 R78-B1 工程单位换算族模板派生首版
 *============================================================================*)
TYPE E_DL_TimeUnit :
(
    eSec := 0,      // 秒 [s] / Second
    eMin,           // 分 [min] / Minute
    eHour           // 时 [h] / Hour
);
END_TYPE

FUNCTION FC_DL_TimeUnitConvert : REAL
VAR_INPUT
    fValue : REAL;         // 输入数值 [源单位] / Input value in source unit
    eSrc : E_DL_TimeUnit;  // 源单位选择 / Source unit selector
    eDst : E_DL_TimeUnit;  // 目标单位选择 / Destination unit selector
END_VAR
VAR
    fBase : REAL;          // 归一化中间值 [s] / Normalized intermediate in seconds
END_VAR
FC_DL_TimeUnitConvert := 0.0;   // 缺省返回 0 / Default return 0
CASE eSrc OF                    // 段 1：归一到基准 s / Normalize to base seconds
    E_DL_TimeUnit.eSec: fBase := fValue;                // 基准直通 / Base pass-through
    E_DL_TimeUnit.eMin: fBase := fValue * 60.0;         // 1 min = 60 s
    E_DL_TimeUnit.eHour: fBase := fValue * 3600.0;      // 1 h = 3600 s
    ELSE FC_DL_TimeUnitConvert := 0.0; RETURN;          // 源枚举非法返 0 / Invalid source returns 0
END_CASE
CASE eDst OF                    // 段 2：基准到目标 / Base to destination
    E_DL_TimeUnit.eSec: FC_DL_TimeUnitConvert := fBase;             // 基准直通 / Base pass-through
    E_DL_TimeUnit.eMin: FC_DL_TimeUnitConvert := fBase / 60.0;      // s 到 min
    E_DL_TimeUnit.eHour: FC_DL_TimeUnitConvert := fBase / 3600.0;   // s 到 h
    ELSE FC_DL_TimeUnitConvert := 0.0;                  // 目标枚举非法返 0 / Invalid destination returns 0
END_CASE
END_FUNCTION

(* ---- FC_DL_TorqueUnitConvert.st ---- *)
//==============================================================================
// 函数：FC_DL_TorqueUnitConvert ｜ 中文名称：转矩单位换算（枚举选路 + 域闸）
// 所属子库：DL_MathData ｜ 版本：v1.0.0 ｜ 日期：2026-11-23
// 兼容：CODESYS V3.5+ / TwinCAT 3 / 汇川 InoProShop / Machine Expert（纯标准库）
// 功能描述：转矩单位双向换算原子：N·m ↔ kgf·m ↔ lb·ft。换算因子取国际
//           公开口径：1 kgf·m = 9.80665 N·m；1 lb·ft = 1.35582 N·m。
//           允许带符号输入（正/负转矩均合法），换算为纯线性乘法。
// 开源溯源 (Origin)：候选队列 MS_TO_KMH（oscatBasic，MIT 许可，
//           https://github.com/tkucic/brOscatLib/blob/main/oscatBasic/MS_TO_KMH.st）
//           ——单位换算族行为定义参考；原名 MS_TO_KMH → 道莅
//           FC_DL_TorqueUnitConvert，clean-room 独立重写（枚举选路 + 域闸
//           增强为道莅防御规范增量，零源码行复制）
// 公开接口清单：输入 eMode / fValue；输出 fResult / bValid
// 错误码表：纯函数无状态机码轨；无效输入经 bValid = FALSE 表达（哨兵返回
//           0.0），本件不占用 16#0001 段码位（邻件免让位）
// 状态机：E_DL_TorqueUnit（本文件唯一定义，全库唯一属主）：
//           eNmToKgm = 0 / eKgmToNm = 1 / eNmToLbFt = 2 / eLbFtToNm = 3；
//           枚举非法值走 CASE ELSE 兜底
// 边界行为：① 任一输入非有限 → 哨兵 0.0 返回；
//           ② 幅值越 LREAL 可表域 → 哨兵 0.0 返回；
//           ③ 枚举非法值 → CASE ELSE 哨兵返回；
//           ④ 纯线性乘法无除法（乘法因子均为常量非零）。
// 修订历史：v1.0.0 2026-11-23 首版（R73 派单 · 批 3 · 序 11）
//==============================================================================

(*------------------------------------------------------------------------------
 * 枚举: E_DL_TorqueUnit（归属本函数，同文件发布，全库唯一属主）
 * 含义: 换算方向选择，成员与 CASE 标签双向完备。
 *-----------------------------------------------------------------------------*)
TYPE E_DL_TorqueUnit :
(
    eNmToKgm  := 0,   // 牛米 → 千克力米 / N·m to kgf·m
    eKgmToNm  := 1,   // 千克力米 → 牛米 / kgf·m to N·m
    eNmToLbFt := 2,   // 牛米 → 磅英尺 / N·m to lb·ft
    eLbFtToNm := 3    // 磅英尺 → 牛米 / lb·ft to N·m
);
END_TYPE

(*------------------------------------------------------------------------------
 * 调用示例：fT := FC_DL_TorqueUnitConvert(
 *             eMode := E_DL_TorqueUnit.eNmToKgm, fValue := 25.0,
 *             bValid => bOk);
 * 注意：仅当 bValid = TRUE 时结果可进入判据；带符号转矩均合法。
 *-----------------------------------------------------------------------------*)
FUNCTION FC_DL_TorqueUnitConvert : LREAL
VAR_INPUT
    eMode    : E_DL_TorqueUnit;        // 换算方向枚举 [—] / Conversion direction enum
    fValue   : LREAL;                  // 输入转矩值 [源单位]，带符号合法 / Torque value [source unit], signed allowed
END_VAR
VAR_OUTPUT
    bValid   : BOOL;                   // 结果有效标志，FALSE 时返回哨兵 0.0 / Result validity flag
END_VAR
VAR CONSTANT
    DL_TQ_KGM  : LREAL := 9.80665;     // 千克力米→牛米因子 [牛米每千克力米] / kgf·m to N·m factor
    DL_TQ_LBFT : LREAL := 1.35582;     // 磅英尺→牛米因子 [牛米每磅英尺] / lb·ft to N·m factor
    DL_TQ_INF  : LREAL := 1.7976931348623157E308; // LREAL 幅值上限 / LREAL magnitude ceiling
    DL_TQ_ZERO : LREAL := 0.0;         // 无效哨兵返回值 / Sentinel return for invalid
END_VAR

// ---- 段 1｜出口默认值（纯函数无实例，无定时器/沿刷新义务）----
bValid := FALSE;                      // 缺省无效 / Invalid by default

// ---- 段 2｜输入防御：非有限值（NaN 自反判 + Inf 幅值判，R79）----
IF (fValue <> fValue) OR (ABS(fValue) > DL_TQ_INF) THEN
    FC_DL_TorqueUnitConvert := DL_TQ_ZERO; // 无效输入：哨兵零返回 / Invalid input, sentinel zero return
    RETURN;                            // 结构早退 / early exit
END_IF

// ---- 段 3｜换算主体（CASE 带 ELSE；纯线性乘法，因子常量非零）----
CASE eMode OF
    E_DL_TorqueUnit.eNmToKgm:          // 牛米 → 千克力米（除以因子，幅值只减不溢）
        FC_DL_TorqueUnitConvert := fValue / DL_TQ_KGM; // 千克力米 [kgf·m] / kgf·m result

    E_DL_TorqueUnit.eKgmToNm:          // 千克力米 → 牛米（乘因子，幅值放大先闸）
        IF ABS(fValue) > (DL_TQ_INF / DL_TQ_KGM) THEN
            FC_DL_TorqueUnitConvert := DL_TQ_ZERO; // 乘积越表域哨兵返回（预检防 Inf 污染）/ Product would overflow, sentinel return
            RETURN;                    // 结构早退 / early exit
        END_IF
        FC_DL_TorqueUnitConvert := fValue * DL_TQ_KGM; // 牛米 [N·m] / N·m result

    E_DL_TorqueUnit.eNmToLbFt:         // 牛米 → 磅英尺（除以因子，幅值只减不溢）
        FC_DL_TorqueUnitConvert := fValue / DL_TQ_LBFT; // 磅英尺 [lb·ft] / lb·ft result

    E_DL_TorqueUnit.eLbFtToNm:         // 磅英尺 → 牛米（乘因子，幅值放大先闸）
        IF ABS(fValue) > (DL_TQ_INF / DL_TQ_LBFT) THEN
            FC_DL_TorqueUnitConvert := DL_TQ_ZERO; // 乘积越表域哨兵返回（预检防 Inf 污染）/ Product would overflow, sentinel return
            RETURN;                    // 结构早退 / early exit
        END_IF
        FC_DL_TorqueUnitConvert := fValue * DL_TQ_LBFT; // 牛米 [N·m] / N·m result

    ELSE                               // 枚举非法值兜底（R21：CASE 必带 ELSE）
        FC_DL_TorqueUnitConvert := DL_TQ_ZERO; // 非法枚举：哨兵零返回 / Illegal enum, sentinel zero return
        RETURN;                        // 结构早退 / early exit
END_CASE

bValid := TRUE;                       // 全部防御通过：结果有效 / Result valid
END_FUNCTION

(* ---- FC_DL_ViscosityUnitConvert.st ---- *)
(*==============================================================================
 * 组件名称 (Component)  : FC_DL_ViscosityUnitConvert
 * 所属子库 (Sublibrary) : DL_MathData
 * 当前版本 (Version)    : 1.0.0
 * 兼容性   (Platform)   : CODESYS 3.5+ / TwinCAT 3 / 汇川 InoProShop / 施耐德 Machine Expert
 *                         仅依赖 IEC 61131-3 算术运算符，零厂商私有库
 * 功能描述 (Function)   : 运动粘度单位换算（系数表驱动）：以 mm²/s 为中介单位，
 *                         fHub = fValue × kSrc，fResult = fHub ÷ kDst；系数为编译期
 *                         非零常量，纯常量除法，结构性无除零。
 *                         **单位恒等说明**：1 cSt ≡ 1 mm²/s（厘斯定义即 mm²/s），
 *                         两成员为同一物理量不同书写，故系数均为 1.0；本件保留两个枚举
 *                         成员以适配不同 HMI 标签与协议字段，避免上游做字符串映射。
 *                         **温度不补偿（适用域声明）**：运动粘度强烈依赖温度，
 *                         本件为纯量纲换算，不引入任何温度修正；调用方必须保证
 *                         参与比较的数据同温基准（推荐 40 ℃ 基准，ISO 3448 VG 体系）。
 *                         粘度非负：负值判故障级 eNegativeValue 并回哨兵 0。
 * 接口     (Interface)  : 输入 fValue 被换算粘度 [源单位]、eSrc 源单位、eDst 目标单位；
 *                         输出 fConverted 换算结果 [目标单位]、eErrCode（E_DL_ViscConvErr）；
 *                         返回值 = bValid 数值可信标志（TRUE = fConverted 可信）。
 * 边界     (Boundary)   : ① 属主边界：只做单位换算，不做温度补偿、不做粘度-温度曲线拟合。
 *                         ② 单位枚举越域 → 故障级 eInvalidUnit，结果哨兵 0。
 *                         ③ 非有限双判，命中即故障级 eNonFinite。
 *                         ④ 负粘度 → 故障级 eNegativeValue（拒绝，不钳位）。
 *                         ⑤ 零粘度 → 信息级 eZeroValue（物理上仅真空/静止，多为未充油）。
 *                         ⑥ m²/s → mm²/s 放大 1E6，结果复检防溢出为非有限。
 *                         ⑦ 零全局耦合（无 GVL / VAR_EXTERNAL / 物理地址）。
 * 分工声明 (Scope)      : 与 `FC_DL_DensityUnitConvert` 分工：密度换算归那件；
 *                         粘度等级（VG32 等）选型属配方管理，不在本件范围。
 * 来源标签 (Source Tag) : 开源溯源：lgf-math 换算系数（公开物理常数，clean-room 重写）；许可证 MIT（仅参考语义，代码原创）
 * 码表     (Codes)      : 本件不占用全局数字码位；出口为 BOOL + LREAL +
 *                         本文件内定义 enum E_DL_ViscConvErr（全库唯一）。
 * 红线自检 (Redline)    : R1 ✓ 零 GVL/VAR_EXTERNAL ｜ R2 ✓ 零 %I/%Q/%M ｜ R3 ✓ 纯 IEC 61131-3
 *                         R4 ✓ 非有限双判 + 枚举域闸 + 常量除法无除零 + 负值拒绝 ｜ R5 ✓ 声明逐行同行双语注释
 *                         R6 N/A（纯函数无状态机） ｜ R7 N/A（无实例调用）
 * 修订历史 (Revision)   : 2026-11-23  v1.0.0  R77 首版（批次 B2 · 序号 16）
 * 验收向量 (Acceptance) : ① fValue=32.0, eSrc=eCst, eDst=eMm2s → 32×1.0 = 32 mm2/s,
 *                         ÷1.0 = 32.0, eOk, TRUE（恒等）；
 *                         ② fValue=1.0, eSrc=eM2s, eDst=eMm2s → 1×1E6 = 1000000.0 mm2/s；
 *                         ③ fValue=1000000.0, eSrc=eMm2s, eDst=eM2s → 1.0 m2/s（容差 1E-12）；
 *                         ④ fValue=-1.0, eSrc=eCst, eDst=eMm2s → 返回 FALSE, 0, eNegativeValue；
 *                         ⑤ fValue=0.0, eSrc=eCst, eDst=eMm2s → 0.0, 返回 TRUE, eZeroValue。
 *==============================================================================*)

(*-----------------------------------------------------------------------------
 * 枚举: E_DL_ViscUnit（运动粘度单位表，归属 DL_MathData，与本件同文件，全库唯一属主）
 *----------------------------------------------------------------------------*)
TYPE E_DL_ViscUnit :
(
    eCst  := 0,   // 厘斯（centi-Stokes，定义上恒等于 mm2/s） / Centistokes, identically equal to mm2/s
    eMm2s := 1,   // 平方毫米每秒（中介单位） / Square millimetre per second, hub unit
    eM2s  := 2    // 平方米每秒（= 1E6 mm2/s） / Square metre per second
);
END_TYPE

(*-----------------------------------------------------------------------------
 * 枚举: E_DL_ViscConvErr（运动粘度换算错误码）
 *----------------------------------------------------------------------------*)
TYPE E_DL_ViscConvErr :
(
    eOk            := 0,   // 信息级：换算完成 / Info: conversion completed
    eZeroValue     := 1,   // 信息级：零粘度（多为未充油） / Info: zero viscosity, often unfilled
    eInvalidUnit   := 2,   // 故障级：单位枚举越域 / Fault: unit enum out of domain
    eNonFinite     := 3,   // 故障级：输入非有限 / Fault: non-finite input
    eNegativeValue := 4    // 故障级：负粘度 / Fault: negative viscosity
);
END_TYPE

FUNCTION FC_DL_ViscosityUnitConvert : BOOL
VAR_INPUT
    fValue : LREAL;          // 被换算运动粘度值 [源单位] / Kinematic viscosity value in source unit
    eSrc   : E_DL_ViscUnit;  // 源单位枚举 [-] / Source unit enum
    eDst   : E_DL_ViscUnit;  // 目标单位枚举 [-] / Destination unit enum
END_VAR
VAR_OUTPUT
    fConverted : LREAL;            // 换算结果 [目标单位] / Converted result
    eErrCode   : E_DL_ViscConvErr; // 错误码出口 [-] / Error code outlet
END_VAR
VAR
    _bNonFin : BOOL;   // 输入非有限当拍标志 [-] / Non-finite input flag
    _fHub    : LREAL;  // 中介粘度值 [mm2/s] / Hub viscosity value in square millimetres per second
END_VAR
VAR CONSTANT
    DL_VIC_CST  : LREAL := 1.0;      // cSt → mm2/s 恒等系数 [-] / Centistokes identity factor
    DL_VIC_MM2S : LREAL := 1.0;      // mm2/s → mm2/s 恒等系数 [-] / Hub identity factor
    DL_VIC_M2S  : LREAL := 1.0E6;    // m2/s → mm2/s 换算系数 [-] / Square metre per second factor
    DL_VIC_ZERO : LREAL := 0.0;      // 零粘度与非有限判零基准 [-] / Zero viscosity and non-finite base
END_VAR

(* —— 段 0：出口预置安全值 —— *)
FC_DL_ViscosityUnitConvert := FALSE;               // 返回值预置无效 / Return preset invalid
fConverted := DL_VIC_ZERO;                         // 结果哨兵 0 / Result sentinel
eErrCode   := E_DL_ViscConvErr.eInvalidUnit;       // 预置最严码 / Preset strictest code

(* —— 段 1：非有限域闸（R79 双判） —— *)
_bNonFin := (fValue <> fValue) OR ((fValue - fValue) <> DL_VIC_ZERO);   // 非有限判定 / Non-finite test
IF _bNonFin THEN
    eErrCode := E_DL_ViscConvErr.eNonFinite;       // 故障级码 / Fault-level code
    RETURN;
END_IF

(* —— 段 2：负粘度域闸 —— *)
IF fValue < DL_VIC_ZERO THEN
    eErrCode := E_DL_ViscConvErr.eNegativeValue;   // 故障级码 / Fault-level code
    RETURN;
END_IF

(* —— 段 3：源单位 → 中介 mm2/s —— *)
IF eSrc = E_DL_ViscUnit.eCst THEN
    _fHub := fValue * DL_VIC_CST;                  // cSt 恒等 / Centistokes identity
ELSIF eSrc = E_DL_ViscUnit.eMm2s THEN
    _fHub := fValue * DL_VIC_MM2S;                 // 直通 / Hub pass-through
ELSIF eSrc = E_DL_ViscUnit.eM2s THEN
    _fHub := fValue * DL_VIC_M2S;                  // m2/s × 1E6 / Square metre per second scaled
ELSE
    RETURN;                                        // 源单位越域 / Source unit out of domain
END_IF

(* —— 段 4：中介 mm2/s → 目标单位（常量除法，分母非零） —— *)
IF eDst = E_DL_ViscUnit.eCst THEN
    fConverted := _fHub / DL_VIC_CST;              // ÷1 恒等 / Divide by identity
ELSIF eDst = E_DL_ViscUnit.eMm2s THEN
    fConverted := _fHub / DL_VIC_MM2S;             // ÷1 / Divide by identity
ELSIF eDst = E_DL_ViscUnit.eM2s THEN
    fConverted := _fHub / DL_VIC_M2S;              // ÷1E6 / Divide by square metre per second factor
ELSE
    eErrCode   := E_DL_ViscConvErr.eInvalidUnit;   // 目标单位越域 / Destination out of domain
    fConverted := DL_VIC_ZERO;
    RETURN;
END_IF

(* —— 段 5：结果非有限复检兜底（1E6 放大后必须复检） —— *)
IF (fConverted <> fConverted) OR ((fConverted - fConverted) <> DL_VIC_ZERO) THEN
    fConverted := DL_VIC_ZERO;                     // 复检异常回哨兵 / Recheck failed: sentinel
    eErrCode   := E_DL_ViscConvErr.eNonFinite;     // 故障级码 / Fault-level code
    RETURN;
END_IF

(* —— 段 6：成功出口 —— *)
IF fValue = DL_VIC_ZERO THEN
    eErrCode := E_DL_ViscConvErr.eZeroValue;       // 信息级：零粘度 / Info: zero viscosity
ELSE
    eErrCode := E_DL_ViscConvErr.eOk;              // 信息级成功 / Info success
END_IF
FC_DL_ViscosityUnitConvert := TRUE;                // 换算有效 / Conversion valid

END_FUNCTION

(* ---- FC_DL_VolumeUnitConvert.st ---- *)
(*==============================================================================
 * 组件名称 (Component)  : FC_DL_VolumeUnitConvert
 * 所属子库 (Sublibrary) : DL_MathData
 * 当前版本 (Version)    : 1.0.0
 * 兼容性   (Platform)   : CODESYS 3.5+ / TwinCAT 3 / 汇川 InoProShop / 施耐德 Machine Expert
 *                         仅依赖 IEC 61131-3 算术运算符，零厂商私有库
 * 功能描述 (Function)   : 体积 / 容积单位换算（系数表驱动）：以升（L）为中介单位，
 *                         fHub = fValue × kSrc，fResult = fHub ÷ kDst；系数为编译期
 *                         非零常量，纯常量除法，结构性无除零。
 *                         体积非负：负值判故障级 eNegativeValue 并回哨兵 0。
 *                         美制加仑采用 US liquid gallon 定义（3.785411784 L），
 *                         与英制加仑（4.54609 L）不同，本件显式标定 US 口径。
 * 接口     (Interface)  : 输入 fValue 被换算体积 [源单位]、eSrc 源单位、eDst 目标单位；
 *                         输出 fConverted 换算结果 [目标单位]、eErrCode（E_DL_VolConvErr）；
 *                         返回值 = bValid 数值可信标志（TRUE = fConverted 可信）。
 * 边界     (Boundary)   : ① 属主边界：只做单位换算，不做罐体液位-体积曲线换算（归查表族）。
 *                         ② 单位枚举越域 → 故障级 eInvalidUnit，结果哨兵 0。
 *                         ③ 非有限双判，命中即故障级 eNonFinite。
 *                         ④ 负体积 → 故障级 eNegativeValue（拒绝，不钳位）。
 *                         ⑤ 零值合法（info 级 eZeroValue）。结果与中介值各复检一次。
 *                         ⑥ **口径声明**：本件 gal 恒为 US liquid gallon = 3.785411784 L。
 *                         ⑦ 零全局耦合（无 GVL / VAR_EXTERNAL / 物理地址）。
 * 分工声明 (Scope)      : 与 `FC_DL_AreaUnitConvert` 分工：面积不做隐式 × 高度推导；
 *                         与 `FC_DL_DensityUnitConvert` 分工：密度归那件，本件不隐含质量。
 * 来源标签 (Source Tag) : 开源溯源：lgf-math 换算系数（公开物理常数，clean-room 重写）；许可证 MIT（仅参考语义，代码原创）
 * 码表     (Codes)      : 本件不占用全局数字码位；出口为 BOOL + LREAL +
 *                         本文件内定义 enum E_DL_VolConvErr（全库唯一）。
 * 红线自检 (Redline)    : R1 ✓ 零 GVL/VAR_EXTERNAL ｜ R2 ✓ 零 %I/%Q/%M ｜ R3 ✓ 纯 IEC 61131-3
 *                         R4 ✓ 非有限双判 + 枚举域闸 + 常量除法无除零 + 负值拒绝 ｜ R5 ✓ 声明逐行同行双语注释
 *                         R6 N/A（纯函数无状态机） ｜ R7 N/A（无实例调用）
 * 修订历史 (Revision)   : 2026-11-23  v1.0.0  R77 首版（批次 B2 · 序号 13）
 * 验收向量 (Acceptance) : ① fValue=1.0, eSrc=eM3, eDst=eL → 1×1000 = 1000.0 L, eOk, TRUE；
 *                         ② fValue=1.0, eSrc=eGalUs, eDst=eL → 3.785411784 L（容差 1E-9）；
 *                         ③ fValue=1000.0, eSrc=eMl, eDst=eL → 1000×0.001 = 1.0 L；
 *                         ④ fValue=-2.0, eSrc=eL, eDst=eMl → 返回 FALSE, 0, eNegativeValue；
 *                         ⑤ fValue=0.0, eSrc=eL, eDst=eM3 → 0.0, 返回 TRUE, eZeroValue。
 *==============================================================================*)

(*-----------------------------------------------------------------------------
 * 枚举: E_DL_VolUnit（体积单位表，归属 DL_MathData，与本件同文件，全库唯一属主）
 *----------------------------------------------------------------------------*)
TYPE E_DL_VolUnit :
(
    eL     := 0,   // 升（中介单位，= 1 dm3） / Litre, hub unit, one cubic decimetre
    eM3    := 1,   // 立方米（1000 L） / Cubic metre, one thousand litres
    eGalUs := 2,   // 美制液量加仑（3.785411784 L） / US liquid gallon
    eMl    := 3    // 毫升（千分之一 L） / Millilitre, one thousandth of litre
);
END_TYPE

(*-----------------------------------------------------------------------------
 * 枚举: E_DL_VolConvErr（体积换算错误码）
 *----------------------------------------------------------------------------*)
TYPE E_DL_VolConvErr :
(
    eOk            := 0,   // 信息级：换算完成 / Info: conversion completed
    eZeroValue     := 1,   // 信息级：输入为零（合法） / Info: zero input, legal
    eInvalidUnit   := 2,   // 故障级：单位枚举越域 / Fault: unit enum out of domain
    eNonFinite     := 3,   // 故障级：输入非有限 / Fault: non-finite input
    eNegativeValue := 4    // 故障级：负体积 / Fault: negative volume
);
END_TYPE

FUNCTION FC_DL_VolumeUnitConvert : BOOL
VAR_INPUT
    fValue : LREAL;          // 被换算体积值 [源单位] / Volume value in source unit
    eSrc   : E_DL_VolUnit;   // 源单位枚举 [-] / Source unit enum
    eDst   : E_DL_VolUnit;   // 目标单位枚举 [-] / Destination unit enum
END_VAR
VAR_OUTPUT
    fConverted : LREAL;           // 换算结果 [目标单位] / Converted result
    eErrCode   : E_DL_VolConvErr; // 错误码出口 [-] / Error code outlet
END_VAR
VAR
    _bNonFin : BOOL;   // 输入非有限当拍标志 [-] / Non-finite input flag
    _fHub    : LREAL;  // 中介体积值 [L] / Hub volume value in litres
END_VAR
VAR CONSTANT
    DL_VUC_L     : LREAL := 1.0;          // L → L 恒等系数 [L/L] / litre identity factor
    DL_VUC_M3    : LREAL := 1000.0;       // m3 → L 换算系数 [L/m3] / cubic metre to litre factor
    DL_VUC_GALUS : LREAL := 3.785411784;  // US gal → L 换算系数 [L/gal] / US gallon to litre factor
    DL_VUC_ML    : LREAL := 0.001;        // mL → L 换算系数 [L/mL] / millilitre to litre factor
    DL_VUC_ZERO  : LREAL := 0.0;          // 零值与非有限判零基准 [-] / Zero and non-finite base
END_VAR

(* —— 段 0：出口预置安全值 —— *)
FC_DL_VolumeUnitConvert := FALSE;                  // 返回值预置无效 / Return preset invalid
fConverted := DL_VUC_ZERO;                         // 结果哨兵 0 / Result sentinel
eErrCode   := E_DL_VolConvErr.eInvalidUnit;        // 预置最严码 / Preset strictest code

(* —— 段 1：非有限域闸（R79 双判） —— *)
_bNonFin := (fValue <> fValue) OR ((fValue - fValue) <> DL_VUC_ZERO);   // 非有限判定 / Non-finite test
IF _bNonFin THEN
    eErrCode := E_DL_VolConvErr.eNonFinite;        // 故障级码 / Fault-level code
    RETURN;
END_IF

(* —— 段 2：负体积域闸 —— *)
IF fValue < DL_VUC_ZERO THEN
    eErrCode := E_DL_VolConvErr.eNegativeValue;    // 故障级码 / Fault-level code
    RETURN;
END_IF

(* —— 段 3：源单位 → 中介升 —— *)
IF eSrc = E_DL_VolUnit.eL THEN
    _fHub := fValue * DL_VUC_L;                    // L 直通 / litre pass-through
ELSIF eSrc = E_DL_VolUnit.eM3 THEN
    _fHub := fValue * DL_VUC_M3;                   // m3 × 1000 / cubic metre scaled
ELSIF eSrc = E_DL_VolUnit.eGalUs THEN
    _fHub := fValue * DL_VUC_GALUS;                // US gal × 3.785411784 / US gallon scaled
ELSIF eSrc = E_DL_VolUnit.eMl THEN
    _fHub := fValue * DL_VUC_ML;                   // mL × 0.001 / millilitre scaled
ELSE
    RETURN;                                        // 源单位越域 / Source unit out of domain
END_IF

(* —— 段 4：中介升 → 目标单位（常量除法，分母非零） —— *)
IF eDst = E_DL_VolUnit.eL THEN
    fConverted := _fHub / DL_VUC_L;                // ÷1 / Divide by identity
ELSIF eDst = E_DL_VolUnit.eM3 THEN
    fConverted := _fHub / DL_VUC_M3;               // ÷1000 / Divide by cubic metre factor
ELSIF eDst = E_DL_VolUnit.eGalUs THEN
    fConverted := _fHub / DL_VUC_GALUS;            // ÷3.785411784 / Divide by US gallon factor
ELSIF eDst = E_DL_VolUnit.eMl THEN
    fConverted := _fHub / DL_VUC_ML;               // ÷0.001 / Divide by millilitre factor
ELSE
    eErrCode   := E_DL_VolConvErr.eInvalidUnit;    // 目标单位越域 / Destination out of domain
    fConverted := DL_VUC_ZERO;
    RETURN;
END_IF

(* —— 段 5：结果非有限复检兜底 —— *)
IF (fConverted <> fConverted) OR ((fConverted - fConverted) <> DL_VUC_ZERO) THEN
    fConverted := DL_VUC_ZERO;                     // 复检异常回哨兵 / Recheck failed: sentinel
    eErrCode   := E_DL_VolConvErr.eNonFinite;      // 故障级码 / Fault-level code
    RETURN;
END_IF

(* —— 段 6：成功出口 —— *)
IF fValue = DL_VUC_ZERO THEN
    eErrCode := E_DL_VolConvErr.eZeroValue;        // 信息级：零值 / Info: zero value
ELSE
    eErrCode := E_DL_VolConvErr.eOk;               // 信息级成功 / Info success
END_IF
FC_DL_VolumeUnitConvert := TRUE;                   // 换算有效 / Conversion valid

END_FUNCTION
